(* IEC 61131-3 sources: daoli-st-library/DL_Process (part 47) *)

(* ---- FB_DL_QuarterCellCutSeq.st ---- *)
(*
  FB_DL_QuarterCellCutSeq  —  极片分切顺控（刀轴相位 + 张力窗 + 废边回收） / Electrode slitting sequencer with blade phase, tension window and trim recovery
  分类 Category : DL_Process
  版本 Version  : 1.0.0
  来源 Source   : roadmap-li-p2 — 锂电极片分切工站真缺口
  溯源 Origin   : 道莅 clean-room 实现；刀轴相位对齐 + 张力窗监督 + 废边回收联锁为公开分切工艺逻辑，未复制任何源码行
  功能 Function : 1) 三段顺控：ePhase 刀轴相位对齐（fBladePhaseDeg 进目标容差带）→
                  eRun 分切运行（张力窗 fTensionN 双向监督 + 废边回收信号 bTrimOk 监督）→
                  eStop 收料停机（tStop 到时）→ eDone；2) 相位对齐超时保护；
                  3) 故障级单码 03A0，归因由 eCause 独立成员承载（R190）；
                  4) 信息级 04C8 = 分切循环完成沿；5) 解除式全当拍量（R240）。
  接口 Interface: 输入相位/张力/废边信号与复位位；输出状态/相位镜像/张力窗镜像/码
  边界 Boundary : ① 组态闸：fPhaseTolDeg <= 0.0、fTensionHiN <= fTensionLoN、tPhaseTmo <= T#0S、
                  tStop <= T#0S → 03A0 锁存；② 相位判据为双向容差式，相位量纲约定
                  0~360 单调注入（跨零归一由调用方完成，本件不内联 MOD 以免非标准扩展）；
                  ③ 浮点禁 = / <> 判等；④ 全部 TON / R_TRIG 段 0 无条件周期调用；
                  ⑤ 故障相迁出唯一路径 = bReset 上升沿；⑥ 零全局耦合（无 GVL / %I %Q %M）。
  依赖 Depends  : Standard.library（TON / R_TRIG）
  码表 Error codes（Process 段 0005，故障窗口 03A0 / 信息窗口 04C8）:
    16#0005_03A0 故障级：分切故障总码（组态非法 / 相位对齐超时 / 张力越窗 / 废边回收异常），
                 锁存至 bReset 上升沿；归因见 eCause，不新增码位（派单硬约束单码）
    16#0005_04C8 信息级：分切循环完成沿（收料停机完成进 eDone 单拍）
  修订历史 Revision :
    2026-11-19  v1.0.0  R43 首版（批次 1 · 序号 4）
*)

TYPE E_DL_QcsState :
(
    eIdle  := 0,      // 未使能待启动 / Idle, waiting start
    ePhase := 10,     // 刀轴相位对齐中 / Blade phase alignment
    eRun   := 20,     // 分切运行（张力窗 + 废边监督） / Slitting under tension and trim supervision
    eStop  := 30,     // 收料停机中 / Web stop
    eDone  := 50,     // 循环完成 / Done
    eFault := 90      // 故障锁存相 / Fault latched phase
);
END_TYPE

TYPE E_DL_QcsCause :
(
    eNone       := 0, // 无故障成因 / No cause
    eCfgIllegal := 1, // 组态非法 / Illegal configuration
    ePhaseTmo   := 2, // 相位对齐超时 / Phase alignment timeout
    eTensionDev := 3, // 张力越窗 / Tension out of window
    eTrimLost   := 4  // 废边回收异常 / Trim recovery lost
);
END_TYPE

FUNCTION_BLOCK FB_DL_QuarterCellCutSeq
VAR_INPUT
    fBladePhaseDeg  : REAL := 0.0;       // 刀轴实测相位 [°]，0~360 单调注入 / Blade shaft phase
    fPhaseTgtDeg    : REAL := 90.0;      // 目标相位 [°] / Target phase
    fPhaseTolDeg    : REAL := 1.0;       // 相位容差带 [°]，域 > 0 / Phase tolerance
    fTensionN       : REAL := 0.0;       // 实测极片张力 [N] / Measured web tension
    fTensionLoN     : REAL := 20.0;      // 张力窗下限 [N] / Tension low limit
    fTensionHiN     : REAL := 60.0;      // 张力窗上限 [N] / Tension high limit
    bTrimOk         : BOOL := FALSE;     // 废边回收正常信号（电平）[-] / Trim recovery healthy
    tPhaseTmo       : TIME := T#5S;      // 相位对齐超时 [ms]，域 > 0 / Phase timeout
    tStop           : TIME := T#2S;      // 收料停机时长 [ms]，域 > 0 / Web stop duration
    bStart          : BOOL := FALSE;     // 启动命令（电平）[-] / Start command
    bReset          : BOOL := FALSE;     // 复位命令，上升沿清故障 [-] / Reset edge
END_VAR
VAR_OUTPUT
    eState          : E_DL_QcsState;     // 状态出口，段 6 单点映射 / State outlet
    eCause          : E_DL_QcsCause;     // 故障成因出口（R190） / Fault cause outlet
    fPhaseDegOut    : REAL;              // 相位镜像 [°] / Phase mirror
    bPhaseOk        : BOOL;              // 相位达窗镜像 [-] / Phase in-window mirror
    bTensionOk      : BOOL;              // 张力在窗镜像 [-] / Tension in-window mirror
    bCycleDone      : BOOL;              // 循环完成标志 [-] / Cycle done flag
    bError          : BOOL;              // 故障锁存标志 [-] / Fault latch flag
    nErrId          : UDINT;             // 事件码，0 = 无事件 / Event code
END_VAR
VAR
    _eState         : E_DL_QcsState := E_DL_QcsState.eIdle;   // 内部相位（CASE 唯一写入目标） / Internal phase
    _eCause         : E_DL_QcsCause := E_DL_QcsCause.eNone;   // 故障成因锁存（锁存量） / Latched cause
    tonPhase        : TON;               // 相位对齐计时，每周期无条件调用 / Phase timer
    tonStop         : TON;               // 收料停机计时，每周期无条件调用 / Stop timer
    rtReset         : R_TRIG;            // 复位沿实例，每周期无条件调用 / Reset edge
    _bPhaseOk       : BOOL;              // 相位达窗当拍量 [-] / Phase verdict
    _bTensionOk     : BOOL;              // 张力在窗当拍量 [-] / Tension verdict
    _bCfgBad        : BOOL;              // 组态非法当拍量 [-] / Config illegal
    _bFault         : BOOL;              // 故障锁存位（锁存量） / Latched fault bit
    _uFault         : UDINT;             // 故障码锁存（锁存量） / Latched fault code
    _uInfo          : UDINT;             // 信息码，每拍重算 / Transient info code
END_VAR

(* —— 段 0：沿实例与定时器无条件周期刷新 —— *)
_bPhaseOk := ABS(fBladePhaseDeg - fPhaseTgtDeg) <= fPhaseTolDeg;                 // 相位容差判据 / Phase tolerance verdict
_bTensionOk := (fTensionN >= fTensionLoN - 1.0E-6) AND (fTensionN <= fTensionHiN + 1.0E-6);  // 张力容差窗 / Tension window verdict
_bCfgBad := (fPhaseTolDeg <= 0.0) OR (fTensionHiN <= fTensionLoN)
            OR (tPhaseTmo <= T#0S) OR (tStop <= T#0S);                          // 组态非法当拍量 / Config illegal
rtReset(CLK := bReset);                                                        // 复位沿，每拍必调 / Reset edge
tonPhase(IN := (_eState = E_DL_QcsState.ePhase), PT := tPhaseTmo);             // 相位对齐计时 / Phase timer
tonStop(IN := (_eState = E_DL_QcsState.eStop), PT := tStop);                   // 收料停机计时 / Stop timer

(* —— 段 1：单拍量预清零（锁存量不入清单） —— *)
_uInfo := 16#0000_0000;            // 信息码每拍重算 / Info recomputed
fPhaseDegOut := 0.0;               // 相位镜像缺省 0 / Phase mirror default
bPhaseOk := FALSE;                 // 相位镜像缺省 FALSE / Phase flag default
bTensionOk := FALSE;               // 张力镜像缺省 FALSE / Tension flag default
bCycleDone := FALSE;               // 完成标志缺省 FALSE / Done default
nErrId := 16#0000_0000;            // 事件码缺省无事件 / Event code default

(* —— 段 2：复位沿 + 组态域闸 —— *)
IF rtReset.Q THEN                              // rtReset.Q = 当拍量 / current scan
    _bFault := FALSE;                          // 清故障锁存位（锁存量） / Clear fault latch
    _uFault := 16#0000_0000;                   // 清故障锁存码（锁存量） / Clear fault code
    _eCause := E_DL_QcsCause.eNone;            // 清成因（锁存量） / Clear cause
    IF _eState = E_DL_QcsState.eFault THEN
        _eState := E_DL_QcsState.eIdle;        // 故障相迁出：回未使能 / Fault exit to idle
    END_IF
END_IF
IF _bCfgBad THEN                               // 组态域闸 / Config gate
    _uFault := 16#0005_03A0;                   // 故障级：分切故障总码 / Process fault code
    _eCause := E_DL_QcsCause.eCfgIllegal;      // 归因：组态非法 / Cause: illegal config
    _bFault := TRUE;                           // 标志与码位配对（R45） / Flag paired with code
END_IF

(* —— 段 3：超时 / 张力越窗 / 废边异常（判据当拍量） —— *)
IF (NOT _bFault) AND tonPhase.Q THEN           // 相位对齐超时 / Phase timeout
    _uFault := 16#0005_03A0;
    _eCause := E_DL_QcsCause.ePhaseTmo;        // 归因：相位超时 / Cause: phase timeout
    _bFault := TRUE;
END_IF
IF (NOT _bFault) AND (_eState = E_DL_QcsState.eRun) AND (NOT _bTensionOk) THEN   // 运行期张力越窗 / Tension deviation
    _uFault := 16#0005_03A0;
    _eCause := E_DL_QcsCause.eTensionDev;      // 归因：张力越窗 / Cause: tension
    _bFault := TRUE;
END_IF
IF (NOT _bFault) AND (_eState = E_DL_QcsState.eRun) AND (NOT bTrimOk) THEN       // 废边回收异常 / Trim lost
    _uFault := 16#0005_03A0;
    _eCause := E_DL_QcsCause.eTrimLost;        // 归因：废边异常 / Cause: trim lost
    _bFault := TRUE;
END_IF

(* —— 段 4：故障解除式（R240；全当拍量）：rtReset.Q / NOT _bCfgBad / NOT tonPhase.Q —— *)
IF rtReset.Q AND (NOT _bCfgBad) AND (NOT tonPhase.Q) THEN
    _bFault := FALSE;                          // 清故障锁存位（锁存量） / Clear fault latch
    _uFault := 16#0000_0000;                   // 清故障锁存码（锁存量） / Clear fault code
    _eCause := E_DL_QcsCause.eNone;            // 清成因（锁存量） / Clear cause
END_IF

(* —— 段 4A：故障锁存相位迁移闸 —— *)
IF _bFault AND (_eState <> E_DL_QcsState.eFault) THEN
    _eState := E_DL_QcsState.eFault;           // 锁存即入故障相 / Latch enters fault phase
END_IF

(* —— 段 5：相位机（CASE 全覆盖 + ELSE 兜底） —— *)
CASE _eState OF

E_DL_QcsState.eIdle:
    IF bStart AND (NOT _bFault) THEN           // 启动条件 / Start gate
        _eState := E_DL_QcsState.ePhase;       // 进相位对齐相 / Enter phase alignment
    END_IF

E_DL_QcsState.ePhase:
    IF _bPhaseOk THEN                          // 出口 1：相位达窗 / Phase reached
        _eState := E_DL_QcsState.eRun;         // 进分切运行相 / Enter slitting
    ELSIF NOT bStart THEN                      // 出口 2：撤启动（R98 双出口） / Start released
        _eState := E_DL_QcsState.eIdle;        // 回未使能 / Back to idle
    END_IF

E_DL_QcsState.eRun:
    IF NOT bStart THEN                         // 撤启动：进停机相 / Start released enters stop
        _eState := E_DL_QcsState.eStop;
    END_IF

E_DL_QcsState.eStop:
    IF tonStop.Q THEN                          // 停机计时到 / Stop elapsed
        _uInfo := 16#0005_04C8;                // 信息级：循环完成沿 / Info: cycle complete edge
        _eState := E_DL_QcsState.eDone;        // 进完成相 / Enter done
    END_IF

E_DL_QcsState.eDone:
    IF bStart THEN                             // 新循环请求 / New cycle request
        _eState := E_DL_QcsState.ePhase;       // 进相位相 / Enter phase
    END_IF

E_DL_QcsState.eFault:
    ;                                          // 故障相：仅段 4 复位沿可迁出 / Only reset exits

ELSE
    _uFault := 16#0005_03A0;                   // 故障级：非法相位兜底（归并总码） / Illegal phase fallback
    _eCause := E_DL_QcsCause.eCfgIllegal;      // 归因：相位非法归并组态 / Cause: phase illegal
    _bFault := TRUE;
    _eState := E_DL_QcsState.eFault;           // 强制回故障相 / Force fault phase

END_CASE

(* —— 段 6：出口单点映射（名实同源；锁存码回放） —— *)
fPhaseDegOut := fBladePhaseDeg;                    // 相位镜像 / Phase mirror
bPhaseOk := _bPhaseOk AND (NOT _bFault);           // 相位达窗镜像 / Phase mirror
bTensionOk := _bTensionOk AND (NOT _bFault);       // 张力窗镜像 / Tension mirror
bCycleDone := (_eState = E_DL_QcsState.eDone);     // 完成标志 / Done flag
IF _bFault THEN
    nErrId := _uFault;                         // 故障锁存码回放 / Replay latched code
ELSE
    nErrId := _uInfo;                          // 信息码 / Transient info
END_IF
bError := _bFault;                             // 故障标志同源 / Flag from latch
eState := _eState;                             // 状态出口 / State outlet
eCause := _eCause;                             // 成因出口 / Cause outlet

END_FUNCTION_BLOCK

(* ---- FB_DL_QuenchTemperLineSeq.st ---- *)
(*==============================================================================
  Component : FB_DL_QuenchTemperLineSeq
  Category  : DL_Process
  Type      : FB
  Complexity: C4
  VERSION   : v1.0.0
  功能      : 淬火-回火联动线全流程顺控（上料/加热/保温/淬火/沥液/回火/冷却/下料）
  开源溯源  : 道莅原创 clean-room 自研（无外部代码引用）｜License: MIT
  边界条件  : ① 本件只编排相与时序闸，不驱动阀门接触器；执行器由 IO 映射层按相指示位驱动。
              ② E1 仅加热相与沥液相可重试（定时器自复位后重新计时），预算 nRetryMax 耗尽升 E2。
              ③ E3 判据（急停断开 / 安全门未闭 / 液位低于下限 / 介质超温）同拍置 bSafeCut；
                 锁存解除唯一路径 = bReset 沿且安全条件已恢复（R152），bStop 不清 E3。
              ④ 配比约束（R100）：atPhaseTmo[1] 加热窗须宽于实测升温时间；atPhaseTmo[6] 回火总窗
                 须 ≥ 升温 + 保温整定之和，否则回火带内判据永不到时。
              ⑤ 复位作用域（R311）：bReset 沿清 E2/E3 锁存 + 节拍累加 + 重试计数；bStop 只清 E2 与相位。
              ⑥ 默认引脚组合自证（R114）：握手类（bPartLoaded / bUnloadPermit / bDrained /
                 bQuenchImmersion）默认 FALSE，默认组合无法越过任一握手直达完成相；使能类（bDoorClosed /
                 bEStopHealthy）默认 TRUE 与 bEnable 同族，断线由硬件安全回路保证，不靠软件默认值兜底。
  状态机    : eIdle 待机 / eLoad 上料 / eHeat 加热 / eSoak 保温 / eQuench 淬火 / eDrain 沥液 /
              eTemper 回火 / eCool 冷却 / eUnload 下料 / eFault 故障停(E2) / eSafeStop 安全断能(E3)
  自检      : R1 零 GVL ｜ R2 零物理地址 ｜ R3 纯 IEC 61131-3 ｜ R4 非有限自反判 + 除零先判 ｜
              R6 CASE 含 ELSE ｜ R7 八 TON 两沿段 0 无条件刷新 ｜ R10 仅标准转换函数 ｜ R14 无属性件
==============================================================================*)
TYPE E_DL_QtlPhase :
(
    eIdle     := 0,     (* 待机：等启动沿 / Idle, waiting for start edge *)
    eLoad     := 10,    (* 上料相：等上料到位 / Loading, wait load-in-position *)
    eHeat     := 20,    (* 加热相：升到保温带（E1 可重试）/ Heating, retryable *)
    eSoak     := 30,    (* 保温相：保温到时 / Soaking *)
    eQuench   := 40,    (* 淬火相：浸没且到时 / Quenching, immersed and timed *)
    eDrain    := 50,    (* 沥液相：等回液到位（E1 可重试）/ Draining, retryable *)
    eTemper   := 60,    (* 回火相：带内且总窗到时 / Tempering, in band and window *)
    eCool     := 70,    (* 冷却相：空冷到出料温度 / Cooling to unload temperature *)
    eUnload   := 80,    (* 下料相：等下料允许 / Unloading, wait permit *)
    eFault    := 90,    (* 故障停待复位（E2）/ Fault stop awaiting reset, E2 *)
    eSafeStop := 95     (* 安全侧断能（E3）/ Safety energy cut, E3 *)
);
END_TYPE
TYPE E_DL_QtlCause :
(
    eNone      := 0,    (* 无异常 / No anomaly *)
    eLoadTmo   := 1,    (* 上料超时 / Load timeout *)
    eHeatTmo   := 2,    (* 加热超时（E1 记录后重试）/ Heat timeout, retried *)
    eSoakTmo   := 3,    (* 保温超时 / Soak timeout *)
    eQuenchTmo := 4,    (* 淬火到时未浸没 / Quench timed out without immersion *)
    eDrainTmo  := 5,    (* 沥液超时（E1 记录后重试）/ Drain timeout, retried *)
    eTemperTmo := 6,    (* 回火超时（带内未达）/ Tempering timeout *)
    eCoolTmo   := 7,    (* 冷却超时 / Cooling timeout *)
    eUnloadTmo := 8,    (* 下料超时 / Unload timeout *)
    eRetryOver := 9,    (* 重试预算耗尽（E1 升 E2）/ Retry budget exhausted *)
    eSigBad    := 10,   (* 工件温度信号非有限（E2）/ Part temperature non-finite *)
    eEstopOpen := 11,   (* 急停回路断开（E3）/ E-stop circuit open *)
    eDoorOpen  := 12,   (* 安全门未闭合（E3）/ Guard door open *)
    eLevelLow  := 13,   (* 淬火槽液位低于下限（E3）/ Bath level low *)
    eMediumHi  := 14,   (* 淬火介质超温（E3）/ Medium over-temperature *)
    eCfgBad    := 15,   (* 组态非法（E2）/ Illegal configuration *)
    ePhaseBad  := 16    (* 非法相位兜底（E2）/ Illegal phase fallback *)
);
END_TYPE
TYPE E_DL_QtlGrade :
(
    eG0 := 0,           (* 无异常 / No anomaly *)
    eG1 := 1,           (* E1 可恢复重试：记录后重试，不置 bError / E1 retried, recorded only *)
    eG2 := 2,           (* E2 停机待复位 / E2 stop, awaiting reset *)
    eG3 := 3            (* E3 安全侧立即断能 / E3 immediate safety energy cut *)
);
END_TYPE

FUNCTION_BLOCK FB_DL_QuenchTemperLineSeq
VAR_INPUT
    bStart        : BOOL := FALSE;      (* 启动沿（eIdle 入 eLoad） [-] / Start rising edge *)
    bStop         : BOOL := FALSE;      (* 中止：回 eIdle 并清 E2 锁存（不清 E3） [-] / Abort, clears E2 only *)
    bReset        : BOOL := FALSE;      (* 复位沿：清全部锁存 + 节拍 + 重试（R311） [-] / Reset edge *)
    bPartLoaded   : BOOL := FALSE;      (* 上料到位（默认 FALSE 禁跳步） [-] / Load in position *)
    bUnloadPermit : BOOL := FALSE;      (* 下料允许（默认 FALSE 禁跳步） [-] / Unload permit *)
    bQuenchOil    : BOOL := TRUE;       (* 介质：TRUE 油淬 / FALSE 水淬 [-] / Oil when TRUE *)
    bQuenchImmersion : BOOL := FALSE;   (* 淬火浸没到位（默认 FALSE 禁跳步） [-] / Quench immersion OK *)
    bDrained      : BOOL := FALSE;      (* 沥液回液到位（默认 FALSE 禁跳步） [-] / Drain back complete *)
    bDoorClosed   : BOOL := TRUE;       (* 安全门闭合（使能类引脚，默认 TRUE） [-] / Guard door closed *)
    bEStopHealthy : BOOL := TRUE;       (* 急停回路正常（使能类引脚，默认 TRUE） [-] / E-stop healthy *)
    fMediumTempC  : LREAL := 0.0;       (* 淬火介质温度实测 [℃] / Medium temperature [degC] *)
    fLevelPct     : LREAL := 0.0;       (* 淬火槽液位实测 [%] / Bath level [%] *)
    fPartTempC    : LREAL := 0.0;       (* 工件温度实测（升温与冷却判据） [℃] / Part temperature [degC] *)
    fSoakSetC     : LREAL := 850.0;     (* 保温设定温度，域 > 0 [℃] / Soak setpoint [degC] *)
    fTemperSetC   : LREAL := 550.0;     (* 回火设定温度，域 > 0 [℃] / Temper setpoint [degC] *)
    fSoakTolC     : LREAL := 15.0;      (* 保温与回火带共用半宽，域 > 0 [℃] / Band half-width [degC] *)
    fMediumMaxC   : LREAL := 60.0;      (* 介质温度上限，域 > 0（E3 判据） [℃] / Medium limit [degC] *)
    fLevelMinPct  : LREAL := 70.0;      (* 液位安全下限，域 0..100（E3 判据） [%] / Level floor [%] *)
    fCoolSetC     : LREAL := 80.0;      (* 冷却出料温度上限，域 > 0 [℃] / Cool-down unload limit [degC] *)
    atPhaseTmo    : ARRAY[0..8] OF TIME := [T#3M, T#45M, T#90M, T#15M, T#8M, T#3M, T#120M, T#30M, T#3M];   (* 超时窗 [ms]，下标 0..8 = 上料/加热/保温/油淬/水淬/沥液/回火/冷却/下料 / Phase windows [ms] *)
    nRetryMax     : UINT := 2;          (* 单相 E1 重试预算，域 1..9（0 入组态闸） [次] / Retry budget *)
    fCycleSec     : LREAL := 0.0;       (* 扫描周期（<=0 用缺省 0.01s） [s] / Scan cycle [s] *)
END_VAR
VAR_OUTPUT
    eState        : E_DL_QtlPhase;      (* 当前相（HMI 诊断） [-] / Present phase *)
    eCause        : E_DL_QtlCause;      (* 成因（锁存回放，R189） [-] / Latched cause playback *)
    eGrade        : E_DL_QtlGrade;      (* 异常分级出口 [-] / Exception grade outlet *)
    bError        : BOOL;               (* 故障标志（E2/E3 为 TRUE，E1 不置） [-] / Error flag *)
    bSafeCut      : BOOL;               (* 安全侧断能指令（E3 常 TRUE 至复位） [-] / Safety energy cut *)
    bHeatActive   : BOOL;               (* 加热相指示（供 IO 层驱动加热阀） [-] / Heating indicator *)
    bQuenchActive : BOOL;               (* 淬火相指示（供 IO 层驱动淬火机构） [-] / Quench indicator *)
    bDone         : BOOL;               (* 单拍完成脉冲 [-] / One-scan done pulse *)
    nPieceCount   : UDINT;              (* 累计产量（饱和于 UDINT 上限） [件] / Piece count, saturating *)
    tCycleLast    : TIME;               (* 最近一件节拍 [ms] / Last piece cycle [ms] *)
    fCycleAvgS    : LREAL;              (* 平均节拍（无件输出 0） [s] / Average cycle [s] *)
    nRetryUsed    : UINT;               (* 当前相已用重试次数 [次] / Retries used in phase *)
END_VAR
VAR
    _ePhase      : E_DL_QtlPhase := E_DL_QtlPhase.eIdle;    (* 内部相（CASE 唯一写入目标） [-] / Internal phase *)
    _ePhasePrev  : E_DL_QtlPhase := E_DL_QtlPhase.eIdle;    (* 上拍相快照（相迁移后置用） [-] / Previous phase *)
    _eCause      : E_DL_QtlCause := E_DL_QtlCause.eNone;    (* 成因锁存量 [-] / Latched cause *)
    _eGrade      : E_DL_QtlGrade := E_DL_QtlGrade.eG0;      (* 分级锁存量 [-] / Latched grade *)
    _bFault      : BOOL := FALSE;       (* E2 锁存位（解除 = bReset 沿或 bStop） [-] / E2 latch *)
    _bSafeLatch  : BOOL := FALSE;       (* E3 锁存位（解除 = bReset 沿且安全恢复） [-] / E3 latch *)
    _bFaultReq   : BOOL := FALSE;       (* 单拍故障请求（段 1 预清，段 6 落地） [-] / One-scan fault request *)
    _bDonePulse  : BOOL := FALSE;       (* 单拍完成标志（段 1 预清） [-] / One-scan done flag *)
    _bMediumBad  : BOOL := FALSE;       (* 介质温度非有限或超上限 [-] / Medium bad *)
    _bLevelBad   : BOOL := FALSE;       (* 液位非有限或低于下限 [-] / Level bad *)
    _bPartBad    : BOOL := FALSE;       (* 工件温度非有限 [-] / Part temperature non-finite *)
    _bSoakBand   : BOOL := FALSE;       (* 保温带内判据 [-] / In soak band *)
    _bTemperBand : BOOL := FALSE;       (* 回火带内判据 [-] / In temper band *)
    _bCfgBad     : BOOL := FALSE;       (* 组态非法当拍量 [-] / Configuration bad *)
    _nRetry      : UINT := 0;           (* 当前相重试计数（相迁移后置清） [次] / Retry counter *)
    _nPiece      : UDINT := 0;          (* 产量累计锁存（饱和） [件] / Piece count latch *)
    _nIdx        : INT := 0;            (* 相窗遍历索引（循环变量） [-] / Loop index *)
    _fCycleAccS  : LREAL := 0.0;        (* 本件节拍累加 [s] / Cycle accumulator *)
    _fCycleSumS  : LREAL := 0.0;        (* 节拍总和（均值分子） [s] / Cycle sum *)
    _fCy         : LREAL := 0.0;        (* 当拍有效周期 [s] / Effective cycle *)
    _tCycleLast  : TIME := T#0S;        (* 最近节拍锁存 [ms] / Last cycle latch *)
    _tQuenchTmo  : TIME := T#15M;       (* 当拍淬火窗（按介质选择） [ms] / Active quench window [ms] *)
    tonLoad      : TON;                 (* 上料超时（段 0 无条件调用） / Load timeout *)
    tonHeat      : TON;                 (* 加热超时（自复位，E1 可重试） / Heat timeout, self-reset *)
    tonSoak      : TON;                 (* 保温超时 / Soak timeout *)
    tonQuench    : TON;                 (* 淬火超时（按介质选窗） / Quench timeout *)
    tonDrain     : TON;                 (* 沥液超时（自复位，E1 可重试） / Drain timeout, self-reset *)
    tonTemper    : TON;                 (* 回火总窗（升温 + 保温） / Temper total window *)
    tonCool      : TON;                 (* 冷却超时 / Cool timeout *)
    tonUnload    : TON;                 (* 下料超时 / Unload timeout *)
    rtStart      : R_TRIG;              (* 启动沿（段 0 无条件调用） / Start edge *)
    rtReset      : R_TRIG;              (* 复位沿（段 0 无条件调用） / Reset edge *)
END_VAR
VAR CONSTANT
    DL_QTL_CYDEF    : LREAL := 0.01;        (* 缺省扫描周期 [s] / Default scan cycle [s] *)
    DL_QTL_PCMAX    : UDINT := 4294967295;  (* 产量计数饱和上限 [件] / Piece count ceiling *)
    DL_QTL_RETRYTOP : UINT := 9;            (* 重试预算可配域顶 [次] / Retry configurable ceiling *)
    DL_QTL_PCTOP    : LREAL := 100.0;       (* 液位百分比满量程 [%] / Level full scale [%] *)
END_VAR

(*-----------------------------------------------------------------------------
  方法 ResetFault：清 E2/E3 锁存（唯一解除入口，R152 可达性自证）
  契约：入参 bSafetyOk 表示安全条件已恢复；返回 TRUE = 本次确实清除了锁存。
  E2 恒可清；E3 仅当 bSafetyOk 为 TRUE 才可清（否则锁存保持，解除路径显式可达）。
  作用域：清 _bFault / _bSafeLatch / _eCause / _eGrade / _nRetry，并把相位迁回 eIdle。
-----------------------------------------------------------------------------*)
METHOD PUBLIC ResetFault : BOOL
VAR_INPUT
    bSafetyOk : BOOL := FALSE;      (* 安全条件已恢复（E3 解除前置） [-] / Safety conditions recovered *)
END_VAR
VAR
    _bCleared : BOOL := FALSE;      (* 本次是否清除过锁存 [-] / Cleared this call *)
END_VAR

ResetFault := FALSE;                (* 返回预置安全值 / Preset safe return *)
_bCleared := FALSE;
IF _bSafeLatch THEN
    IF bSafetyOk THEN
        _bSafeLatch := FALSE;       (* E3 解除：安全侧恢复后允许 / E3 released after safety recovery *)
        _bCleared := TRUE;
    END_IF
ELSIF _bFault THEN
    _bFault := FALSE;               (* E2 解除：无条件可清 / E2 released unconditionally *)
    _bCleared := TRUE;
END_IF
IF _bCleared THEN
    _eCause := E_DL_QtlCause.eNone;     (* 清成因 / Clear cause *)
    _eGrade := E_DL_QtlGrade.eG0;       (* 清分级 / Clear grade *)
    _nRetry := 0;                       (* 清重试预算占用 / Clear retry usage *)
    _ePhase := E_DL_QtlPhase.eIdle;     (* 迁回待机 / Back to idle *)
END_IF
ResetFault := _bCleared;            (* 真值返回 / Final return *)
END_METHOD

(*-----------------------------------------------------------------------------
  方法 CalcCycleTime：本件节拍换算（毫秒取整 + 双向域闸，无跨周期驻留）
  口径：NaN 自反检出 -> 返回哨兵零点 T#0S（还原方向不饱和，R81）；
        Inf 用差值自减检出 -> 亦返回哨兵零点；负值拒收；
        超 TIME 可表上限先钳后转（R153 取整前实数上限兜底）。
-----------------------------------------------------------------------------*)
METHOD PUBLIC CalcCycleTime : TIME
VAR
    fMs   : LREAL := 0.0;           (* 节拍毫秒暂存 [ms] / Milliseconds scratch *)
    fMsCl : LREAL := 0.0;           (* 钳位后毫秒 [ms] / Clamped milliseconds *)
    diMs  : DINT := 0;              (* 整型毫秒（钳位后转换，防溢出翻转） [ms] / Integer milliseconds *)
END_VAR

CalcCycleTime := T#0S;              (* 哨兵零点 / Sentinel zero *)
fMs := _fCycleAccS * 1000.0;        (* 秒 -> 毫秒 [ms] / Second to millisecond *)
IF (fMs <> fMs) OR ((fMs - fMs) <> (fMs - fMs)) OR (fMs < 0.0) THEN
    CalcCycleTime := T#0S;          (* 域闸：NaN 自反 / Inf 差值自减 / 负值，均拒收 / Domain gate *)
    RETURN;
END_IF
IF fMs > 2147483647.0 THEN
    fMsCl := 2147483647.0;          (* 先钳到 TIME 可表毫秒上限 / Clamp to TIME ceiling *)
ELSE
    fMsCl := fMs;
END_IF
diMs := LREAL_TO_DINT(fMsCl);       (* 钳位后整型转换（R10 标准函数） / Clamped integer conversion *)
CalcCycleTime := DINT_TO_TIME(diMs);(* 标准转换链 / Standard conversion chain *)
END_METHOD

(* —— 段 0：三模拟量非有限判定 + 组态闸 + 淬火窗选择 + 周期派生 + 八 TON 两沿无条件刷新（R7） —— *)
_bMediumBad := (fMediumTempC <> fMediumTempC)
            OR ((fMediumTempC - fMediumTempC) <> (fMediumTempC - fMediumTempC))
            OR (fMediumTempC > fMediumMaxC);      (* NaN 自反 + Inf 差值 + 超上限 / NaN, Inf, over-limit *)
_bLevelBad := (fLevelPct <> fLevelPct)
           OR ((fLevelPct - fLevelPct) <> (fLevelPct - fLevelPct))
           OR (fLevelPct < fLevelMinPct);         (* NaN 自反 + Inf 差值 + 低于下限 / NaN, Inf, low level *)
_bPartBad := (fPartTempC <> fPartTempC)
          OR ((fPartTempC - fPartTempC) <> (fPartTempC - fPartTempC));   (* 工件温度非有限 / Part temp non-finite *)
_bCfgBad := (nRetryMax = 0) OR (nRetryMax > DL_QTL_RETRYTOP)
         OR (fSoakSetC <= 0.0) OR (fTemperSetC <= 0.0) OR (fSoakTolC <= 0.0)
         OR (fMediumMaxC <= 0.0) OR (fCoolSetC <= 0.0)
         OR (fLevelMinPct < 0.0) OR (fLevelMinPct > DL_QTL_PCTOP);   (* 静态组态域闸全枚举 / Static config gate *)
FOR _nIdx := 0 TO 8 DO
    IF atPhaseTmo[_nIdx] <= T#0S THEN
        _bCfgBad := TRUE;                          (* 任一相窗非正 -> 组态非法 / Non-positive phase window *)
    END_IF
END_FOR
IF bQuenchOil THEN
    _tQuenchTmo := atPhaseTmo[3];                  (* 油淬窗 / Oil quench window *)
ELSE
    _tQuenchTmo := atPhaseTmo[4];                  (* 水淬窗 / Water quench window *)
END_IF
IF fCycleSec > 0.0 THEN
    _fCy := fCycleSec;                             (* 组态周期有效 / Configured cycle valid *)
ELSE
    _fCy := DL_QTL_CYDEF;                          (* 周期缺省兜底 / Default cycle *)
END_IF
_bSoakBand := (NOT _bPartBad) AND (ABS(fPartTempC - fSoakSetC) <= fSoakTolC);     (* 保温带内（容差比较） / In soak band *)
_bTemperBand := (NOT _bPartBad) AND (ABS(fPartTempC - fTemperSetC) <= fSoakTolC); (* 回火带内（共用半宽） / In temper band *)
rtStart(CLK := bStart);                            (* 启动沿，每拍必调 / Start edge every scan *)
rtReset(CLK := bReset);                            (* 复位沿，每拍必调 / Reset edge every scan *)
tonLoad(IN := (_ePhase = E_DL_QtlPhase.eLoad), PT := atPhaseTmo[0]);              (* 上料超时 / Load window *)
tonHeat(IN := (_ePhase = E_DL_QtlPhase.eHeat) AND (NOT tonHeat.Q), PT := atPhaseTmo[1]);   (* 加热自复位窗（R188） / Heat self-reset *)
tonSoak(IN := (_ePhase = E_DL_QtlPhase.eSoak), PT := atPhaseTmo[2]);              (* 保温超时 / Soak window *)
tonQuench(IN := (_ePhase = E_DL_QtlPhase.eQuench), PT := _tQuenchTmo);            (* 淬火超时 / Quench window *)
tonDrain(IN := (_ePhase = E_DL_QtlPhase.eDrain) AND (NOT tonDrain.Q), PT := atPhaseTmo[5]); (* 沥液自复位窗 / Drain self-reset *)
tonTemper(IN := (_ePhase = E_DL_QtlPhase.eTemper), PT := atPhaseTmo[6]);          (* 回火总窗 / Temper window *)
tonCool(IN := (_ePhase = E_DL_QtlPhase.eCool), PT := atPhaseTmo[7]);              (* 冷却超时 / Cool window *)
tonUnload(IN := (_ePhase = E_DL_QtlPhase.eUnload), PT := atPhaseTmo[8]);          (* 下料超时 / Unload window *)

(* —— 段 1：单拍量预清零（不含锁存/累加/快照量，R107）+ 相迁移后置 —— *)
_bFaultReq := FALSE;                               (* 单拍故障请求预清 / Fault request preset *)
_bDonePulse := FALSE;                              (* 单拍完成标志预清 / Done pulse preset *)
bError := FALSE;                                   (* 故障标志预清（出口 OR 汇总） / Error preset *)
IF _ePhase <> _ePhasePrev THEN
    _nRetry := 0;                                  (* 相迁移：重试预算复位 / Phase change: retry reset *)
    IF _eGrade = E_DL_QtlGrade.eG1 THEN
        _eGrade := E_DL_QtlGrade.eG0;              (* E1 记录随相推进清零（信息级可重算） / E1 cleared on advance *)
        _eCause := E_DL_QtlCause.eNone;
    END_IF
END_IF

(* —— 段 2：E3 安全侧拦截（最高优先级，同拍断能 + 归因唯一 + 迁相） —— *)
IF (NOT bEStopHealthy) OR (NOT bDoorClosed) OR _bLevelBad OR _bMediumBad THEN
    IF NOT _bSafeLatch THEN
        _bSafeLatch := TRUE;                       (* 锁存 / Latch *)
        _eGrade := E_DL_QtlGrade.eG3;              (* 分级 E3 / Grade E3 *)
        bError := TRUE;                            (* 分级标志同段置位（R45 配对） / Error pairing *)
        IF NOT bEStopHealthy THEN
            _eCause := E_DL_QtlCause.eEstopOpen;   (* 归因：急停断开 / Cause: E-stop *)
        ELSIF NOT bDoorClosed THEN
            _eCause := E_DL_QtlCause.eDoorOpen;    (* 归因：安全门未闭 / Cause: door *)
        ELSIF _bLevelBad THEN
            _eCause := E_DL_QtlCause.eLevelLow;    (* 归因：液位低 / Cause: level *)
        ELSE
            _eCause := E_DL_QtlCause.eMediumHi;    (* 归因：介质超温 / Cause: medium *)
        END_IF
    END_IF
    _ePhase := E_DL_QtlPhase.eSafeStop;            (* 同步迁安全相 / Migrate to safety stop *)
END_IF

(* —— 段 3：组态闸入 E2（E3 优先，安全相内不重复置因） —— *)
IF _bCfgBad AND (NOT _bSafeLatch) AND (NOT _bFault) THEN
    _bFault := TRUE;                               (* E2 锁存 / Latch E2 *)
    _eGrade := E_DL_QtlGrade.eG2;                  (* 分级 E2 / Grade E2 *)
    _eCause := E_DL_QtlCause.eCfgBad;              (* 归因：组态非法 / Cause: config *)
    _ePhase := E_DL_QtlPhase.eFault;               (* 同步迁相（R252） / Migrate *)
END_IF

(* —— 段 4：迁出链（复位沿 > 中止；作用域逐项声明 R311） —— *)
IF rtReset.Q THEN
    _bFault := FALSE;                              (* 作用域①：清 E2 锁存 / Clear E2 *)
    IF NOT ((NOT bEStopHealthy) OR (NOT bDoorClosed) OR _bLevelBad OR _bMediumBad) THEN
        _bSafeLatch := FALSE;                      (* 作用域②：安全恢复才清 E3 / Clear E3 only if safe *)
    END_IF
    _eCause := E_DL_QtlCause.eNone;                (* 作用域③：清成因与分级 / Clear cause and grade *)
    _eGrade := E_DL_QtlGrade.eG0;
    _nRetry := 0;                                  (* 作用域④：清重试 / Clear retry *)
    _fCycleAccS := 0.0;                            (* 作用域⑤：清本件节拍累加 / Clear cycle accumulator *)
    IF NOT _bSafeLatch THEN
        IF (_ePhase = E_DL_QtlPhase.eFault) OR (_ePhase = E_DL_QtlPhase.eSafeStop) THEN
            _ePhase := E_DL_QtlPhase.eIdle;        (* 作用域⑥：故障相迁回待机 / Back to idle *)
        END_IF
    END_IF
ELSIF bStop AND (_ePhase <> E_DL_QtlPhase.eIdle) AND (_ePhase <> E_DL_QtlPhase.eSafeStop) THEN
    IF _ePhase = E_DL_QtlPhase.eFault THEN
        _bFault := FALSE;                          (* 中止清 E2（E3 只能由复位清） / Abort clears E2 only *)
        _eCause := E_DL_QtlCause.eNone;
        _eGrade := E_DL_QtlGrade.eG0;
    END_IF
    _nRetry := 0;                                  (* 重试复位 / Retry reset *)
    _fCycleAccS := 0.0;                            (* 节拍累加作废 / Cycle accumulator void *)
    _ePhase := E_DL_QtlPhase.eIdle;                (* 回待机 / Back to idle *)
END_IF

(* —— 段 5：本件节拍累加（仅工作相计时，故障与安全相不累） —— *)
IF (_ePhase <> E_DL_QtlPhase.eIdle) AND (_ePhase <> E_DL_QtlPhase.eFault) AND (_ePhase <> E_DL_QtlPhase.eSafeStop) THEN
    _fCycleAccS := _fCycleAccS + _fCy;
END_IF

(* —— 段 6：故障请求统一落地（分支内只写成因与请求，落地仅此一处，R187/R252） —— *)
IF _bFaultReq AND (NOT _bSafeLatch) THEN
    _bFault := TRUE;                               (* E2 锁存 / Latch E2 *)
    _eGrade := E_DL_QtlGrade.eG2;                  (* 分级 E2 / Grade E2 *)
    _ePhase := E_DL_QtlPhase.eFault;               (* 同步迁相（R252） / Migrate *)
    bError := TRUE;                                (* 故障标志同段置位（R45 配对） / Error pairing *)
END_IF

(* —— 段 7：主状态机（ENUM + CASE，ELSE 兜底回安全相） —— *)
CASE _ePhase OF
E_DL_QtlPhase.eIdle:
    IF rtStart.Q AND (NOT _bFault) AND (NOT _bSafeLatch) THEN
        _fCycleAccS := 0.0;                        (* 新件起算 / New piece *)
        _ePhase := E_DL_QtlPhase.eLoad;            (* 入上料相 / To loading *)
    END_IF
E_DL_QtlPhase.eLoad:
    IF bPartLoaded THEN
        _ePhase := E_DL_QtlPhase.eHeat;            (* 上料到位 -> 加热 / Loaded, heat *)
    ELSIF tonLoad.Q THEN
        _eCause := E_DL_QtlCause.eLoadTmo;         (* 归因：上料超时 / Cause: load timeout *)
        _bFaultReq := TRUE;
    END_IF
E_DL_QtlPhase.eHeat:
    IF _bPartBad THEN
        _eCause := E_DL_QtlCause.eSigBad;          (* 归因：温度信号非有限 / Cause: signal *)
        _bFaultReq := TRUE;
    ELSIF _bSoakBand THEN
        _ePhase := E_DL_QtlPhase.eSoak;            (* 到保温带 -> 保温 / In band, soak *)
    ELSIF tonHeat.Q THEN
        IF _nRetry < nRetryMax THEN
            _nRetry := _nRetry + 1;                (* E1：可重试，计时器自复位后重计时 / E1 retry *)
            _eGrade := E_DL_QtlGrade.eG1;
            _eCause := E_DL_QtlCause.eHeatTmo;
        ELSE
            _eCause := E_DL_QtlCause.eRetryOver;   (* 归因：重试耗尽 / Cause: retry exhausted *)
            _bFaultReq := TRUE;
        END_IF
    END_IF
E_DL_QtlPhase.eSoak:
    IF tonSoak.Q AND _bSoakBand THEN
        _ePhase := E_DL_QtlPhase.eQuench;          (* 到时且带内 -> 淬火 / Timed and in band, quench *)
    ELSIF tonSoak.Q THEN
        _eCause := E_DL_QtlCause.eSoakTmo;         (* 归因：到时仍带外 / Cause: out of band at timeout *)
        _bFaultReq := TRUE;
    END_IF
E_DL_QtlPhase.eQuench:
    IF tonQuench.Q AND bQuenchImmersion THEN
        _ePhase := E_DL_QtlPhase.eDrain;           (* 浸没到位且到时 -> 沥液 / Immersed and timed *)
    ELSIF tonQuench.Q THEN
        _eCause := E_DL_QtlCause.eQuenchTmo;       (* 归因：到时未浸没 / Cause: not immersed *)
        _bFaultReq := TRUE;
    END_IF
E_DL_QtlPhase.eDrain:
    IF bDrained THEN
        _ePhase := E_DL_QtlPhase.eTemper;          (* 回液到位 -> 回火 / Drained, temper *)
    ELSIF tonDrain.Q THEN
        IF _nRetry < nRetryMax THEN
            _nRetry := _nRetry + 1;                (* E1：可重试 / E1 retry *)
            _eGrade := E_DL_QtlGrade.eG1;
            _eCause := E_DL_QtlCause.eDrainTmo;
        ELSE
            _eCause := E_DL_QtlCause.eRetryOver;   (* 归因：重试耗尽 / Cause: retry exhausted *)
            _bFaultReq := TRUE;
        END_IF
    END_IF
E_DL_QtlPhase.eTemper:
    IF _bTemperBand AND tonTemper.Q THEN
        _ePhase := E_DL_QtlPhase.eCool;            (* 带内且总窗到 -> 冷却 / In band and window done *)
    ELSIF tonTemper.Q THEN
        _eCause := E_DL_QtlCause.eTemperTmo;       (* 归因：回火超时（带内未达） / Cause: temper timeout *)
        _bFaultReq := TRUE;
    END_IF
E_DL_QtlPhase.eCool:
    IF _bPartBad THEN
        _eCause := E_DL_QtlCause.eSigBad;          (* 归因：温度信号非有限 / Cause: signal *)
        _bFaultReq := TRUE;
    ELSIF fPartTempC <= fCoolSetC THEN
        _ePhase := E_DL_QtlPhase.eUnload;          (* 冷到出料温度 -> 下料 / Cooled, unload *)
    ELSIF tonCool.Q THEN
        _eCause := E_DL_QtlCause.eCoolTmo;         (* 归因：冷却超时 / Cause: cool timeout *)
        _bFaultReq := TRUE;
    END_IF
E_DL_QtlPhase.eUnload:
    IF bUnloadPermit THEN
        _bDonePulse := TRUE;                       (* 单拍完成（段 1 预清） / One-scan done *)
        _tCycleLast := CalcCycleTime();            (* 委托方法换算节拍 / Delegate cycle conversion *)
        _fCycleSumS := _fCycleSumS + _fCycleAccS;  (* 节拍总和累加 / Cycle sum *)
        _fCycleAccS := 0.0;                        (* 本件累加清零 / Clear accumulator *)
        IF _nPiece < DL_QTL_PCMAX THEN
            _nPiece := _nPiece + 1;                (* 产量推进（容量载体判上限） / Saturating count *)
        END_IF
        _ePhase := E_DL_QtlPhase.eIdle;            (* 回待机迎下一件 / Back to idle *)
    ELSIF tonUnload.Q THEN
        _eCause := E_DL_QtlCause.eUnloadTmo;       (* 归因：下料超时 / Cause: unload timeout *)
        _bFaultReq := TRUE;
    END_IF
E_DL_QtlPhase.eFault:
    bError := TRUE;                                (* 故障相驻留（锁存回放） / Fault residency *)
E_DL_QtlPhase.eSafeStop:
    bError := TRUE;                                (* 安全相驻留（锁存回放） / Safety residency *)
ELSE
    _eCause := E_DL_QtlCause.ePhaseBad;            (* 非法相位兜底 / Illegal phase fallback *)
    _bFault := TRUE;                               (* 兜底锁存 / Fallback latch *)
    _eGrade := E_DL_QtlGrade.eG2;                  (* 兜底分级 E2 / Fallback grade *)
    _ePhase := E_DL_QtlPhase.eFault;               (* 回安全侧 / Fall back to fault *)
    bError := TRUE;
END_CASE

(* —— 段 8：统一出口（电平量由 _ePhase 派生，单拍量由 _b* 标志映射） —— *)
eState := _ePhase;                                 (* 相出口 / Phase outlet *)
eCause := _eCause;                                 (* 成因回放 / Cause playback *)
eGrade := _eGrade;                                 (* 分级出口 / Grade outlet *)
bError := bError OR _bFault OR _bSafeLatch;        (* 故障标志汇总（E1 不置） / Error summary *)
bSafeCut := _bSafeLatch;                           (* 安全断能指令 / Safety energy cut *)
bHeatActive := (_ePhase = E_DL_QtlPhase.eHeat);    (* 加热相指示 / Heating indicator *)
bQuenchActive := (_ePhase = E_DL_QtlPhase.eQuench);(* 淬火相指示 / Quench indicator *)
bDone := _bDonePulse;                              (* 单拍完成脉冲 / One-scan done *)
nPieceCount := _nPiece;                            (* 产量出口 / Count outlet *)
tCycleLast := _tCycleLast;                         (* 节拍出口 [ms] / Cycle outlet *)
IF _nPiece > 0 THEN
    fCycleAvgS := _fCycleSumS / UDINT_TO_LREAL(_nPiece);   (* 均值分母已判非零 / Guarded mean *)
ELSE
    fCycleAvgS := 0.0;                             (* 无件输出 0 / No piece, zero *)
END_IF
nRetryUsed := _nRetry;                             (* 重试占用出口 / Retry outlet *)
_ePhasePrev := _ePhase;                            (* 段末相快照（下拍迁移后置用） / Phase snapshot *)
END_FUNCTION_BLOCK

(* ---- FB_DL_RadiatorZoneValve.st ---- *)
(*
  FB_DL_RadiatorZoneValve  —  散热器末端温控阀脉冲控制 / Radiator zone valve pulse control
  分类 Category : DL_Process
  码位 Code     : 16#06_0_B9
  段位说明      : R38 W7 预留 B6~BF 本轮正式启用，B8 格由 CartonDenestPush 启用，本件启用 B9 格
  版本 Version  : 1.0.0
  来源 Source   : t2-2-lbp — FB_DL_ThreePointValve 典型消费场景待挖项
  溯源 Origin   : clean-room 实现，三点浮阀 + 房间温度闭环为公开经典控制语义，未复制任何源码行
  功能 Function : 1) 房间温度闭环：FC_DL_Hysteresis 迟滞判热需求（fRoomSpC 设定 + fBandC 回差带，
                  带内保持，防阀频繁切换）；
                  2) FB_DL_ThreePointValve 实例消费：热需求 → 开阀指令，无需求 → 关阀指令；
                  3) 最小启停间隔保护：全开后 tMinRun 内禁关、全关后 tMinOff 内禁开
                  （tonMinRun/tonMinOff 双实例，被闭锁期间置信息级码）；
                  4) 阀门限位开关与行程时间由组态透传，估算开度镜像出口。
  边界 Boundary : ① 本件只出三点阀开关指令（经 FB_DL_ThreePointValve 输出脉冲），不写物理 IO；
                  ② 温度信号非有限：需求冻结保持（不误开不误关）+ 信息级码；
                  ③ R228-A 达标声明：tonMinRun/tonMinOff 各自单用途计时（IN 为单相等式），
                  无跨相复用问题（本件无状态机相）；
                  ④ 组态域闸覆盖全部参与换算引脚（R151）；迟滞带/间隔域非法判组态错锁存；
                  ⑤ 需求判据取反口径：迟滞件 TRUE = 温度高（停热），需求 = NOT 迟滞输出，
                  上电冷态需求为 TRUE（保守供热侧）。
  依赖 Depends  : FB_DL_ThreePointValve（实例化，引脚按 registry 实名）；
                  FC_DL_Hysteresis（函数调用，bState 由本件成员持有回传）
  码表 Error codes（本件格 06_0_B9，子码步进 +0x100）:
    16#0006_01B9 信息级：最小启停间隔闭锁中（指令暂缓，不置故障）
    16#0006_02B9 故障级：组态非法（设定/回差/间隔域非法），锁存至复位
    16#0006_03B9 信息级：温度信号非有限，需求冻结保持
    16#0006_04B9 信息级：加热需求置位（bHeating 拍）
    16#0006_05B9 故障级：保留码，本件无 CASE 主状态机，仅作后续维护者新增分支时的防御式默认码

  修订历史 Revision :
    2026-11-19  v1.0.0  R39 首版（批次 4 · 序号 17）
*)

FUNCTION_BLOCK FB_DL_RadiatorZoneValve
VAR_INPUT
    bEnable      : BOOL := TRUE;       // 总使能，FALSE 时关阀指令并冻结需求 [-] / Master enable
    fRoomTempC   : REAL := 20.0;       // 房间实测温度 [°C] / Room measured temperature
    fRoomSpC     : REAL := 21.0;       // 房间设定温度 [°C] / Room setpoint
    fBandC       : REAL := 0.5;        // 需求回差带 [°C]，域 > 0 / Demand hysteresis band
    bLimOpen     : BOOL := FALSE;      // 阀全开限位反馈（透传三点阀）[-] / Valve open limit, passed through
    bLimClosed   : BOOL := FALSE;      // 阀全关限位反馈（透传三点阀）[-] / Valve closed limit, passed through
    tStrokeOpen  : TIME := T#60S;      // 全行程开启时间 [ms]（透传三点阀）/ Full-open stroke time
    tStrokeClose : TIME := T#60S;      // 全行程关闭时间 [ms]（透传三点阀）/ Full-close stroke time
    tMinRun      : TIME := T#120S;     // 最小运行间隔（全开后禁关时长）[ms]，域 >= 0 / Minimum run time
    tMinOff      : TIME := T#120S;     // 最小停歇间隔（全关后禁开时长）[ms]，域 >= 0 / Minimum off time
    bReset       : BOOL := FALSE;      // 故障复位，上升沿生效 / Fault reset, rising edge
END_VAR
VAR_OUTPUT
    bHeating     : BOOL;               // 加热需求（迟滞后，电平）[-] / Heating demand, level
    bOpenCmd     : BOOL;               // 开阀指令生效中（透传阀件脉冲前）[-] / Open command active
    bCloseCmd    : BOOL;               // 关阀指令生效中 [-] / Close command active
    bOpened      : BOOL;               // 阀全开确认（限位优先）[-] / Valve fully opened
    bClosed      : BOOL;               // 阀全关确认（限位优先）[-] / Valve fully closed
    fValvePosEst : REAL;               // 阀估算开度 [%]（三点阀积分口径）/ Valve estimated position
    bError       : BOOL;               // 故障锁存，仅故障级码置位，bReset 清除 [-] / Fault latch
    uErrorId     : UDINT;              // 事件码，0 = 无事件（故障级锁存回放）/ Event code
END_VAR
VAR
    fbValve    : FB_DL_ThreePointValve;   // 三点浮阀实例（主体首部无条件刷新）/ Three-point valve instance
    tonMinRun  : TON;                     // 最小运行计时（全开期间，单用途）/ Minimum run timer, single purpose
    tonMinOff  : TON;                     // 最小停歇计时（全关期间，单用途）/ Minimum off timer, single purpose
    rtReset    : R_TRIG;                  // 复位上升沿 / Reset rising edge
    _bTempHigh : BOOL;                    // 迟滞判温高回传保持变量 / Hysteresis temp-high hold member
    _bHeatDem  : BOOL := TRUE;            // 热需求内部量（上电冷态为 TRUE，保守供热）/ Internal heat demand, TRUE on cold start
    _bTempBad  : BOOL;                    // 温度非有限标志 / Temperature non-finite flag
    _bOpenReq  : BOOL;                    // 开阀请求（需求 + 间隔闭锁裁决后）/ Open request after gating
    _bCloseReq : BOOL;                    // 关阀请求（需求取反 + 间隔闭锁裁决后）/ Close request after gating
    _bBlocked  : BOOL;                    // 本拍指令被间隔闭锁标志 / Command blocked by interval this cycle
    _bOpenedPrv: BOOL;                    // 上拍全开确认镜像（间隔计时基准）/ Previous fully-open mirror, timer basis
    _bClosedPrv: BOOL;                    // 上拍全关确认镜像（间隔计时基准）/ Previous fully-closed mirror, timer basis
    _uInfo     : UDINT;                   // 信息码，每拍重算 / Info code
    _uFault    : UDINT;                   // 故障码锁存寄存 / Latched fault code register
    _bFault    : BOOL;                    // 故障锁存位 / Latched fault bit
    _bCfgBad   : BOOL;                    // 组态非法聚合 / Configuration invalid aggregate
END_VAR
VAR CONSTANT
    DL_RZV_INF_CAP : REAL := 1.0E15;  // 非有限值筛查幅值上限 / Non-finite screening cap
END_VAR

(* —— 段 0：定时器与边沿实例无条件周期刷新（R182：调用语句不得置于 IF/CASE 内） —— *)
(* 间隔计时 IN 取上拍阀位确认镜像（SemaMutex 同款「IN 取上一拍锁存状态」口径） *)
rtReset(CLK := bReset);                                 // 复位沿刷新，每拍必调
tonMinRun(IN := _bOpenedPrv, PT := tMinRun);            // 最小运行计时（上拍全开电平，单用途）
tonMinOff(IN := _bClosedPrv, PT := tMinOff);            // 最小停歇计时（上拍全关电平，单用途）

(* —— 段 1：单拍量预清零（锁存量 _uFault/_bFault/_bHeatDem/_bTempHigh 不入清单，R187①） —— *)
_uInfo := 16#0000_0000;             // 信息码每拍重算
_bCfgBad := FALSE;                  // 组态非法预清零
_bBlocked := FALSE;                 // 闭锁标志预清零
uErrorId := 16#0000_0000;           // 事件码缺省无事件

(* —— 段 3：组态域闸（覆盖全部参与判据换算的引脚，R151） —— *)
IF (fRoomTempC <> fRoomTempC) OR (ABS(fRoomTempC) > DL_RZV_INF_CAP) OR ((fRoomTempC - fRoomTempC) <> 0.0)
   OR (fRoomSpC <> fRoomSpC) OR (ABS(fRoomSpC) > DL_RZV_INF_CAP) THEN
    _bTempBad := TRUE;              // 温度/设定非有限（需求冻结保持，信息级）
END_IF
IF (fBandC <= 0.0) OR (TIME_TO_DINT(tMinRun) < 0) OR (TIME_TO_DINT(tMinOff) < 0)
   OR (TIME_TO_DINT(tStrokeOpen) <= 0) OR (TIME_TO_DINT(tStrokeClose) <= 0) THEN
    _bCfgBad := TRUE;               // 回差/间隔/行程域非法
END_IF
IF _bCfgBad AND (NOT _bFault) THEN
    _uFault := 16#0006_02B9;        // 故障级：组态非法（仅首次进入时写入）
    _bFault := TRUE;
END_IF
IF rtReset.Q AND (NOT _bCfgBad) THEN
    _bFault := FALSE;               // 清故障锁存位（R228-B：rtReset.Q 恒可达）
    _uFault := 16#0000_0000;
END_IF

(* —— 段 4：需求判定（迟滞取反口径；非有限冻结保持） —— *)
IF (NOT _bTempBad) AND (NOT _bCfgBad) THEN
    _bTempHigh := FC_DL_Hysteresis(fIn := fRoomTempC,       // 迟滞判温高（TRUE = 停热侧）
                                   fThreshold := fRoomSpC,  // 设定点
                                   fHysteresis := fBandC,   // 回差带
                                   bState := _bTempHigh);   // 回传保持变量（同一成员，有状态纪律）
    _bHeatDem := NOT _bTempHigh;    // 需求 = NOT 温高（带内保持，防阀频切）
    IF _bHeatDem THEN
        _uInfo := 16#0006_01B9;     // 信息级：加热需求置位
    END_IF
ELSE
    _uInfo := 16#0006_03B9;         // 信息级：温度信号非有限，需求冻结保持（_bHeatDem 不改写）
END_IF

(* —— 段 5：最小启停间隔裁决（先于三点阀调用，数据流「先算后喂」） —— *)
IF NOT bEnable THEN
    _bOpenReq := FALSE;             // 失能：禁开
    _bCloseReq := TRUE;             // 失能：关阀（安全供热侧）
    _bHeatDem := FALSE;             // 失能：需求清零（出口同步）
ELSIF _bFault THEN
    _bOpenReq := FALSE;             // 故障：禁开
    _bCloseReq := TRUE;             // 故障：关阀（安全侧）
    _bHeatDem := FALSE;             // 故障：需求清零（出口同步）
ELSE
    _bOpenReq := _bHeatDem AND (NOT tonMinOff.Q);   // 开阀 = 需求 AND 非停歇闭锁
    _bCloseReq := (NOT _bHeatDem) AND (NOT tonMinRun.Q);    // 关阀 = 无需求 AND 非运行闭锁
    IF _bHeatDem AND tonMinOff.Q THEN
        _bBlocked := TRUE;          // 开阀被停歇闭锁
    END_IF
    IF (NOT _bHeatDem) AND tonMinRun.Q THEN
        _bBlocked := TRUE;          // 关阀被运行闭锁
    END_IF
END_IF
IF _bBlocked THEN
    _uInfo := 16#0006_01B9;         // 信息级：间隔闭锁中（覆盖需求码，闭锁状态优先）
END_IF

(* —— 段 6：三点阀实例调用（每拍顶层无条件；裁决结果作引脚） —— *)
fbValve(bCmdOpen := _bOpenReq,      // 开阀指令（电平）
        bCmdClose := _bCloseReq,    // 关阀指令（电平；与开同拍为假，裁决互斥）
        bLimOpen := bLimOpen,       // 限位透传
        bLimClosed := bLimClosed,   // 限位透传
        tStrokeOpen := tStrokeOpen, // 行程透传
        tStrokeClose := tStrokeClose,   // 行程透传
        fEstimateTol := 10.0,       // 估算-限位一致性容差（默认口径）
        bEnable := TRUE,            // 阀件动作联锁恒放行（闭锁已在本件裁决）
        bReset := bReset,           // 复位透传
        bTrack := FALSE);           // 不跟踪（限位开关口径由透传承载）

(* —— 段 7：出口单点映射（名实同源；锁存码回放，禁同拍抹除） —— *)
_bOpenedPrv := fbValve.bOpened;     // 上拍全开镜像更新（下一拍间隔计时基准）
_bClosedPrv := fbValve.bClosed;     // 上拍全关镜像更新
bHeating := _bHeatDem;              // 需求出口镜像
bOpenCmd := fbValve.bOpenPulse;     // 开阀脉冲镜像（阀件输出）
bCloseCmd := fbValve.bClosePulse;   // 关阀脉冲镜像
bOpened := fbValve.bOpened;         // 全开确认镜像
bClosed := fbValve.bClosed;         // 全关确认镜像
fValvePosEst := fbValve.fPosEstimate;   // 估算开度镜像
IF _bFault THEN
    uErrorId := _uFault;            // 故障锁存码回放
    bError := TRUE;
ELSE
    uErrorId := _uInfo;             // 信息码
    bError := FALSE;
END_IF

END_FUNCTION_BLOCK

(* ---- FB_DL_ReactorChargeSeq.st ---- *)
(*
  DL Factory R84 | FB_DL_ReactorChargeSeq
  功能：反应釜多组分投料顺序时序，逐相流量累积达标判据与搅拌运行互锁
  开源溯源：无（clean-room 自研，依据公开工艺公式，来源=行业通用公式，许可证=MIT，借鉴点=公式结构）
  规则：R1-R16 全遵守
*)
TYPE E_DL_RctChgState :
(
    eIdle := 0, // 空闲待启动 [-] / idle [-]
    eStirCheck := 1, // 搅拌运行确认相 [-] / stirrer check phase [-]
    eChargeA := 2, // A 组分投料相 [-] / component A charging phase [-]
    eChargeB := 3, // B 组分投料相 [-] / component B charging phase [-]
    eChargeC := 4, // C 组分投料相 [-] / component C charging phase [-]
    eHold := 5, // 投料后保持相 [-] / post charge hold phase [-]
    eDone := 6, // 完成相 [-] / done phase [-]
    eFault := 7 // 故障锁存相 [-] / fault latched phase [-]
) := eIdle;
END_TYPE

FUNCTION_BLOCK FB_DL_ReactorChargeSeq
VAR_INPUT
    xStart : BOOL; // 投料启动按钮 [-] / charge start pushbutton [-]
    xReset : BOOL; // 复位按钮，上升沿清故障码与累积量 [-] / reset pushbutton [-]
    xStirRunning : BOOL; // 搅拌运行反馈（投料互锁条件） [-] / stirrer running interlock feedback [-]
    fFlowKgh : REAL; // 当前投料瞬时流量 [kg/h] / instantaneous charge flow [kg/h]
    tScan : TIME := T#50MS; // 扫描周期（累积用） [s] / scan period for accumulation [s]
    aTargetKg : ARRAY[0..2] OF REAL; // A/B/C 三组分目标投料量 [kg] / target mass per component [kg]
    tStirLimit : TIME := T#10S; // 搅拌确认超时 [s] / stirrer check timeout [s]
    tPhaseLimit : TIME := T#600S; // 单组分投料相超时 [s] / per component charge timeout [s]
    tHoldLimit : TIME := T#120S; // 投料后保持时长 [s] / post charge hold duration [s]
END_VAR
VAR_OUTPUT
    eState : E_DL_RctChgState; // 当前时序状态 [-] / current sequence state [-]
    iErrCode : INT; // 故障码 0=正常，501~506 [-] / error code, 501 to 506 [code]
    fChargedKg : REAL; // 本批已投料累计质量 [kg] / total charged mass of this batch [kg]
    xDone : BOOL; // 完成单拍脉冲 [-] / done one-shot pulse [-]
END_VAR
VAR
    rtStart : R_TRIG; // 启动上升沿实例 [-] / start rising edge instance [-]
    rtReset : R_TRIG; // 复位上升沿实例 [-] / reset edge instance [-]
    tonStir : TON; // 搅拌确认超时定时器 [-] / stirrer check timer [-]
    tonPhaseA : TON; // A 组分投料超时定时器（各相独立，R571） [-] / component A charge timer, one per phase [-]
    tonPhaseB : TON; // B 组分投料超时定时器（各相独立，R571） [-] / component B charge timer, one per phase [-]
    tonPhaseC : TON; // C 组分投料超时定时器（各相独立，R571） [-] / component C charge timer, one per phase [-]
    tonHold : TON; // 保持相定时器 [-] / hold phase timer [-]
    _eState : E_DL_RctChgState := E_DL_RctChgState.eIdle; // 内部相位（CASE 唯一写目标） [-] / internal phase [-]
    _iErr : INT; // 故障码内部锁存 [-] / latched error code [-]
    fCharged : REAL; // 累计投料量内部量 [kg] / internal charged mass [kg]
    fPhaseKg : REAL; // 当前组分已投量 [kg] / mass charged in the current phase [kg]
    fDtSec : REAL; // 扫描周期秒值 [s] / scan period in seconds [s]
    fStepKg : REAL; // 本拍投料增量 [kg] / charge increment of this scan [kg]
    xDoneInt : BOOL; // 完成内部锁存位 [-] / internal done latch [-]
    xDonePrev : BOOL; // 完成前拍快照 [-] / done previous scan snapshot [-]
END_VAR

// 段 0｜边沿与定时器实例无条件周期刷新（R7）
rtStart(CLK := xStart); // 启动沿每拍必调 [-] / start edge every scan [-]
rtReset(CLK := xReset); // 复位沿每拍必调 [-] / reset edge every scan [-]
tonStir(IN := _eState = E_DL_RctChgState.eStirCheck, PT := tStirLimit); // 搅拌确认相闸 [-] / stirrer check phase gate [-]
tonPhaseA(IN := _eState = E_DL_RctChgState.eChargeA, PT := tPhaseLimit); // A 相独立计时，离相即复位 [-] / component A timer, reset when the phase leaves [-]
tonPhaseB(IN := _eState = E_DL_RctChgState.eChargeB, PT := tPhaseLimit); // B 相独立计时，离相即复位 [-] / component B timer, reset when the phase leaves [-]
tonPhaseC(IN := _eState = E_DL_RctChgState.eChargeC, PT := tPhaseLimit); // C 相独立计时，离相即复位 [-] / component C timer, reset when the phase leaves [-]
tonHold(IN := _eState = E_DL_RctChgState.eHold, PT := tHoldLimit); // 保持相闸 [-] / hold phase gate [-]

// 段 1｜本拍增量派生（kg/h × s ÷ 3600 = kg）
fDtSec := LREAL_TO_REAL(TIME_TO_LREAL(tScan) / 1000.0); // ms ÷ 1000 = s / [ms] / 1000 = [s]
fStepKg := 0.0; // 增量初值零 [kg] / increment starts at zero [kg]
IF (fFlowKgh > -1.0E30 AND fFlowKgh < 1.0E30) AND fFlowKgh > 0.0 THEN
    fStepKg := (fFlowKgh * fDtSec) / 3600.0; // kg/h × s ÷ 3600 s/h = kg / [kg/h] × [s] / 3600 = [kg]
END_IF

// 段 2｜复位沿：清故障码、累积量与相位（R189）
IF rtReset.Q THEN
    _iErr := 0; // 清故障码 [-] / clear error code [-]
    fCharged := 0.0; // 清本批累计投料 [kg] / clear the batch charge [kg]
    fPhaseKg := 0.0; // 清当前组分累计 [kg] / clear the phase charge [kg]
    xDoneInt := FALSE; // 清完成锁存 [-] / clear done latch [-]
    _eState := E_DL_RctChgState.eIdle; // 回空闲相 [-] / back to idle [-]
END_IF

// 段 3｜主状态机（合法事件优先于超时迁移，R275）
CASE _eState OF
    E_DL_RctChgState.eIdle: // 空闲相 [-] / idle [-]
        xDoneInt := FALSE; // 空闲清完成锁存 [-] / clear done latch in idle [-]
        fCharged := 0.0; // 空闲期累计归零 [kg] / hold the accumulator at zero [kg]
        fPhaseKg := 0.0; // 空闲期组分累计归零 [kg] / hold the phase accumulator at zero [kg]
        IF rtStart.Q THEN
            _eState := E_DL_RctChgState.eStirCheck; // 启动沿先确认搅拌 [-] / start edge checks the stirrer [-]
        END_IF
    E_DL_RctChgState.eStirCheck: // 搅拌确认相（互锁：未运行禁投料） [-] / stirrer check [-]
        IF xStirRunning AND NOT tonStir.Q THEN
            _eState := E_DL_RctChgState.eChargeA; // 搅拌运行转 A 组分 [-] / stirrer running leads to component A [-]
        ELSIF tonStir.Q THEN
            _iErr := 501; _eState := E_DL_RctChgState.eFault; // 搅拌未运行超时（禁投料） [-] / stirrer timeout, charging blocked [-]
        END_IF
    E_DL_RctChgState.eChargeA: // A 组分投料相 [-] / component A [-]
        IF NOT xStirRunning THEN
            _iErr := 502; _eState := E_DL_RctChgState.eFault; // 投料中搅拌停转（互锁断开） [-] / stirrer lost during charging [-]
        ELSIF fPhaseKg >= aTargetKg[0] THEN
            fPhaseKg := 0.0; // 本组分累计清零 [kg] / clear the phase accumulator [kg]
            _eState := E_DL_RctChgState.eChargeB; // A 达标转 B [-] / A reached leads to B [-]
        ELSIF tonPhaseA.Q THEN
            _iErr := 503; _eState := E_DL_RctChgState.eFault; // A 组分投料超时 [-] / component A timeout [-]
        ELSE
            fCharged := fCharged + fStepKg; // kg + kg = kg / [kg] + [kg] = [kg]
            fPhaseKg := fPhaseKg + fStepKg; // kg + kg = kg / [kg] + [kg] = [kg]
        END_IF
    E_DL_RctChgState.eChargeB: // B 组分投料相 [-] / component B [-]
        IF NOT xStirRunning THEN
            _iErr := 502; _eState := E_DL_RctChgState.eFault; // 投料中搅拌停转 [-] / stirrer lost during charging [-]
        ELSIF fPhaseKg >= aTargetKg[1] THEN
            fPhaseKg := 0.0; // 本组分累计清零 [kg] / clear the phase accumulator [kg]
            _eState := E_DL_RctChgState.eChargeC; // B 达标转 C [-] / B reached leads to C [-]
        ELSIF tonPhaseB.Q THEN
            _iErr := 504; _eState := E_DL_RctChgState.eFault; // B 组分投料超时 [-] / component B timeout [-]
        ELSE
            fCharged := fCharged + fStepKg; // kg + kg = kg / [kg] + [kg] = [kg]
            fPhaseKg := fPhaseKg + fStepKg; // kg + kg = kg / [kg] + [kg] = [kg]
        END_IF
    E_DL_RctChgState.eChargeC: // C 组分投料相 [-] / component C [-]
        IF NOT xStirRunning THEN
            _iErr := 502; _eState := E_DL_RctChgState.eFault; // 投料中搅拌停转 [-] / stirrer lost during charging [-]
        ELSIF fPhaseKg >= aTargetKg[2] THEN
            fPhaseKg := 0.0; // 本组分累计清零 [kg] / clear the phase accumulator [kg]
            _eState := E_DL_RctChgState.eHold; // C 达标转保持相 [-] / C reached leads to hold [-]
        ELSIF tonPhaseC.Q THEN
            _iErr := 505; _eState := E_DL_RctChgState.eFault; // C 组分投料超时 [-] / component C timeout [-]
        ELSE
            fCharged := fCharged + fStepKg; // kg + kg = kg / [kg] + [kg] = [kg]
            fPhaseKg := fPhaseKg + fStepKg; // kg + kg = kg / [kg] + [kg] = [kg]
        END_IF
    E_DL_RctChgState.eHold: // 保持相：搅拌必须仍在运行 [-] / hold phase [-]
        IF NOT xStirRunning THEN
            _iErr := 502; _eState := E_DL_RctChgState.eFault; // 保持期搅拌停转 [-] / stirrer lost during hold [-]
        ELSIF tonHold.Q THEN
            _eState := E_DL_RctChgState.eDone; // 保持时长到转完成相 [-] / hold done leads to done [-]
        END_IF
    E_DL_RctChgState.eDone: // 完成相 [-] / done [-]
        xDoneInt := TRUE; // 置完成锁存（出口统一映射单拍） [-] / raise done latch [-]
        IF NOT xStart THEN
            _eState := E_DL_RctChgState.eIdle; // 松开启动即回空闲 [-] / start released returns to idle [-]
        END_IF
    E_DL_RctChgState.eFault: // 故障相：码值锁存回放，仅复位沿出 [-] / fault, exit only on reset [-]
        ; // 锁存回放（R28） [-] / replay the latch only [-]
ELSE
    _iErr := 506; _eState := E_DL_RctChgState.eFault; // 非法相位兜底 [-] / illegal phase fallback [-]
END_CASE

// 段 4｜出口映射（名实双出口，同源赋值）
eState := _eState; // 状态出口 [-] / state outlet [-]
iErrCode := _iErr; // 故障码出口（锁存值） [-] / error code outlet [-]
fChargedKg := fCharged; // 累计投料出口 [kg] / charged mass outlet [kg]
xDone := xDoneInt AND NOT xDonePrev; // 完成单拍（内部锁存 → 出口映射） [-] / done one-shot [-]
xDonePrev := xDoneInt; // 本拍快照供下拍比较 [-] / snapshot for the next scan [-]
END_FUNCTION_BLOCK

(* ---- FB_DL_ReactorRunawayGuard.st ---- *)
(*
  DL Factory R84 | FB_DL_ReactorRunawayGuard
  功能：间歇反应釜放热失控五级联锁：温升速率、绝热温升外推 MTSR、冷却能力失效三判据并行分档，合成 0~5 级动作需求；升级立即生效、降级按延时逐级回落，五级动作位互斥且可降级；L5 全停锁存至复位沿。
  开源溯源：无（clean-room 自研，依据公开工艺公式与安全设计惯例，来源=行业通用公式+工程实践，许可证=MIT，借鉴点=公式结构与联锁分层）
  规则：R1-R16 全遵守
  ------------------------------------------------------------------
  分类 DL_Process ｜ 复杂度 cx5 ｜ 版本 v1.0.0 ｜ 平台 纯 IEC 61131-3（TON、R_TRIG、LREAL、ENUM、CASE）
  边界一：只出分级动作位与诊断量，不驱动泄放阀、冷却阀与投料阀本体，不采集变送器（属主边界，执行由下层 PRG 完成）。
  边界二：三判据分档——判据①温升速率按 fRateTripKmin 的 0.50/0.65/0.80/0.92/1.00 五档；判据②MTSR 按安全裕度 fMtsrMarginK 的已耗比例 0.50/0.35/0.20/0.08/0.00 五档；
          判据③冷却能力按流量下限与夹套-进水温差反向分 3 档与 4 档，温差反向且流量低于半限时直接判 5 档。
  边界三：MTSR 公式＝反应温度 ＋ 累积投料若全部反应的绝热温升：ΔTad [K]＝|ΔH| [kJ/mol] × 1000 [mol/kmol] × 累积摩尔数 [kmol] ÷（批量 [kg] × cp [kJ/(kg·K)]），
          累积摩尔数 [kmol]＝累积投料 [kg] ÷ 平均摩尔质量 [kg/kmol]；ΔTad 上限兜底 300 K 防外推发散。
  边界四：平均摩尔质量 DL_RAG_MOLAR_KGKMOL 为物料体系代理常量——代理值是反应主料的平均摩尔质量、覆盖 100~200 g/mol 的常规精细化工体系、
          体系外（聚合/无机盐）由上层以实测绝热温升标定后换算入参负责（R95 三句齐备，代理假设挂编译验证债）。
  边界五：分级互斥与可降级——iStage 为唯一权威（0~5 整数），五级位按 xStageN＝(iStage ≥ N) 单源派生；升级无延时（安全侧优先），
          降级由 tDegrade 周期窗逐级回落，窗为自复位形式（IN 串 NOT 自身 Q，R188），故不存在同拍双窗，R100 配比约束不适用（本件只有一件定时器）。
  边界六：相位由分级单源映射、零滞后（R191 名实同源），不设独立相位状态机与分级机双权威。
  安全侧：任一浮点入参非有限、组态越域、或任一判据达 5 档 → 立即迁 eTrip 并锁存 xTripLatched；锁存唯一解除路径为 bReset 上升沿（R188），其余路径（失能、条件消失）均不解锁。
  码表：故障级 2711 入参非有限、2712 组态越域、2713 温升速率达 5 档、2714 MTSR 达 5 档、2715 冷却完全失效、2716 非法分级值（防御性保留）；
        以上六码锁存回放且置 bError（R45 配对）；信息级 2701~2705＝当前分级（1~5 级）之动作码，每拍重算且不置 bError。
  输出契约：xStage1..xStage5 为累积电平（N 级生效则 1..N 位全真，互斥性由 iStage 单源保证）；xAlarmOut/xFeedStop/xMaxCool/xVentCmd/xTotalStop 与分级同源派生；
          fMtsrC/fRateKmin/fDtAdK 为诊断连续量，非有限时出零不外抛；xValid 在锁存或闸不过时为假。
  修订记录：2026-11-24 v1.0.0 R84 首版（批 R84 · 序号 42）
*)

TYPE E_DL_RagState :
(
    eNormal   := 0, // 正常：零级，无动作 / normal, level zero, no action
    eWarn     := 1, // 报警：一级，仅告知 / warn, level one, notification only
    eStopFeed := 2, // 停止投料：二级 / stop feeding, level two
    eMaxCool  := 3, // 加大冷却：三级 / maximum cooling, level three
    eVent     := 4, // 紧急泄放：四级 / emergency venting, level four
    eTrip     := 5  // 全停：五级，锁存至复位沿 / total trip, level five, latched until the reset edge
);
END_TYPE

TYPE E_DL_RagCause :
(
    eNone      := 0, // 无成因 / no cause
    eNotFinite := 1, // 入参非有限（故障级 2711）/ a non-finite input, fault grade 2711
    eCfgBad    := 2, // 组态越域（故障级 2712）/ the configuration is out of its domain, fault grade 2712
    eRateHigh  := 3, // 温升速率达五档（故障级 2713）/ the temperature rate reached level five, fault grade 2713
    eMtsrHigh  := 4, // MTSR 达五档（故障级 2714）/ the MTSR reached level five, fault grade 2714
    eCoolLoss  := 5, // 冷却完全失效（故障级 2715）/ the cooling capability was lost, fault grade 2715
    eStageBad  := 6  // 非法分级值（故障级 2716，防御性保留）/ an illegal stage value, fault grade 2716
);
END_TYPE

FUNCTION_BLOCK FB_DL_ReactorRunawayGuard
VAR CONSTANT
    DL_RAG_SEC_MIN     : LREAL := 60.0;    // 秒到分钟折算系数 [s/min] / the second to minute factor [s/min]
    DL_RAG_DT_MIN      : LREAL := 0.001;   // 采样周期下限（速率分母零闸）[s] / the sample period lower bound [s]
    DL_RAG_RATE_ALPHA  : LREAL := 0.30;    // 速率一阶滤波系数 [-] / the first order gain of the rate filter [-]
    DL_RAG_L1_FRAC     : LREAL := 0.50;    // 判据①一级档位系数（跳闸速率的倍数）[-] / the level one factor of the rate criterion [-]
    DL_RAG_L2_FRAC     : LREAL := 0.65;    // 判据①二级档位系数 [-] / the level two factor of the rate criterion [-]
    DL_RAG_L3_FRAC     : LREAL := 0.80;    // 判据①三级档位系数 [-] / the level three factor of the rate criterion [-]
    DL_RAG_L4_FRAC     : LREAL := 0.92;    // 判据①四级档位系数 [-] / the level four factor of the rate criterion [-]
    DL_RAG_M1_FRAC     : LREAL := 0.50;    // 判据②一级档位（裕度已耗比例）[-] / the level one factor of the MTSR criterion [-]
    DL_RAG_M2_FRAC     : LREAL := 0.35;    // 判据②二级档位 [-] / the level two factor of the MTSR criterion [-]
    DL_RAG_M3_FRAC     : LREAL := 0.20;    // 判据②三级档位 [-] / the level three factor of the MTSR criterion [-]
    DL_RAG_M4_FRAC     : LREAL := 0.08;    // 判据②四级档位 [-] / the level four factor of the MTSR criterion [-]
    DL_RAG_COOL_DT_MIN : LREAL := 2.0;     // 夹套与进水温差下限（低于即冷却不足）[K] / the jacket to inlet temperature difference floor [K]
    DL_RAG_FLOW_L4_FRAC: LREAL := 0.50;    // 判据③四级档位流量系数（下限倍数）[-] / the level four flow factor of the cooling criterion [-]
    DL_RAG_DTAD_MAX    : LREAL := 300.0;   // 绝热温升外推上限兜底 [K] / the adiabatic rise extrapolation upper clamp [K]
    DL_RAG_FRAC_MAX    : LREAL := 1.50;    // 已投料占比上限（外推兜底）[-] / the charged fraction upper clamp [-]
    DL_RAG_MOLAR_KGKMOL: LREAL := 100.0;   // 平均摩尔质量代理常量 [kg/kmol] / the mean molar mass proxy [kg/kmol]
    DL_RAG_MOL_PER_KMOL: LREAL := 1000.0;  // 摩尔到千摩尔折算系数 [mol/kmol] / the mole to kilomole factor [mol/kmol]
    DL_RAG_EPS         : LREAL := 1.0E-9;  // 除法零闸与零判定门限 [-] / the division guard and zero test threshold [-]
END_VAR
VAR_INPUT
    bEnable      : BOOL := TRUE;     // 使能，失能只回零级不解除锁存 [-] / enable, a disable only clears the stage and never the latch
    bReset       : BOOL := FALSE;   // 复位上升沿清全停锁存（唯一解除路径）[-] / reset rising edge clears the trip latch, the only release path
    xStirRun     : BOOL := TRUE;    // 搅拌运行反馈，停搅即二级以上 [-] / the agitator running feedback, a stop forces level two or higher
    fTreactC     : LREAL := 25.0;   // 反应温度 [°C] / the reaction temperature [°C]
    fTjacketC    : LREAL := 25.0;   // 夹套温度 [°C] / the jacket temperature [°C]
    fCoolFlowM3h : LREAL := 10.0;   // 冷却水流量 [m³/h] / the cooling water flow [m3/h]
    fCoolInC     : LREAL := 20.0;   // 冷却水进水温度 [°C] / the cooling water inlet temperature [°C]
    fAccumKg     : LREAL := 0.0;    // 累积投料质量（尚未反应部分）[kg] / the accumulated charged mass still unreacted [kg]
    fBatchKg     : LREAL := 1000.0; // 批量总质量 [kg] / the total batch mass [kg]
    fDhKjMol     : LREAL := 80.0;   // 反应焓变（取绝对值参与外推）[kJ/mol] / the reaction enthalpy, the absolute value is used [kJ/mol]
    fCpKjKgK     : LREAL := 3.50;   // 反应液比热容 [kJ/(kg·K)] / the reaction mixture specific heat [kJ/(kg*K)]
    fRateTripKmin: LREAL := 3.00;   // 温升速率跳闸值（五档基准）[K/min] / the rate trip value, the level five base [K/min]
    fMtsrLimitC  : LREAL := 180.0;  // MTSR 安全极限温度 [°C] / the MTSR safety limit temperature [°C]
    fMtsrMarginK : LREAL := 20.0;   // MTSR 安全裕度（分级带宽）[K] / the MTSR safety margin, the staging band [K]
    fFlowMinM3h  : LREAL := 4.00;   // 冷却水流量下限 [m³/h] / the cooling water flow floor [m3/h]
    fDtSec       : LREAL := 0.10;   // 温度采样周期（速率分母）[s] / the temperature sample period, the rate denominator [s]
    tDegrade     : TIME := T#30S;   // 分级降级延时（逐级回落窗）[毫秒] / the stage downgrade delay per step [ms]
END_VAR
VAR_OUTPUT
    eState       : E_DL_RagState := E_DL_RagState.eNormal; // 相位出口（由分级单源映射）[枚举] / the phase outlet mapped from the stage [enum]
    iStage       : INT := 0;      // 当前动作级（0~5，唯一权威）[级] / the active stage, the single authority [level]
    iErrCode     : INT := 0;      // 错误码（故障级锁存回放，信息级每拍重算）[码] / the error code, latched faults and scan info [code]
    bError       : BOOL := FALSE; // 故障标志（与故障级码同源）[-] / the fault flag sharing the fault code source
    xTripLatched : BOOL := FALSE; // 全停锁存（仅复位沿清除）[-] / the trip latch, cleared by the reset edge only
    xValid       : BOOL := FALSE; // 本拍输入与组态可信 [-] / the inputs and the configuration are trustworthy
    xStage1      : BOOL := FALSE; // 一级动作位：报警 [-] / level one action, the alarm
    xStage2      : BOOL := FALSE; // 二级动作位：停止投料 [-] / level two action, stop the feed
    xStage3      : BOOL := FALSE; // 三级动作位：加大冷却 [-] / level three action, maximum cooling
    xStage4      : BOOL := FALSE; // 四级动作位：紧急泄放 [-] / level four action, emergency venting
    xStage5      : BOOL := FALSE; // 五级动作位：全停 [-] / level five action, total trip
    xAlarmOut    : BOOL := FALSE; // 报警输出（一级及以上）[-] / the alarm output from level one on
    xFeedStop    : BOOL := FALSE; // 停止投料输出（二级及以上）[-] / the feed stop output from level two on
    xMaxCool     : BOOL := FALSE; // 加大冷却输出（三级及以上）[-] / the maximum cooling output from level three on
    xVentCmd     : BOOL := FALSE; // 紧急泄放输出（四级及以上）[-] / the emergency vent output from level four on
    xTotalStop   : BOOL := FALSE; // 全停输出（五级）[-] / the total stop output at level five
    fMtsrC       : LREAL := 0.0;  // MTSR 外推值 [°C] / the extrapolated MTSR [°C]
    fRateKmin    : LREAL := 0.0;  // 滤波后温升速率 [K/min] / the filtered temperature rise rate [K/min]
    fDtAdK       : LREAL := 0.0;  // 绝热温升外推量 [K] / the adiabatic rise extrapolation [K]
END_VAR
VAR
    rtReset    : R_TRIG; // 复位沿实例（无量纲）[-] / the reset edge refreshed unconditionally
    tonDown    : TON;    // 降级窗实例（无量纲）[-] / the self resetting downgrade window, its own output inverted
    _eState    : E_DL_RagState := E_DL_RagState.eNormal; // 内部相位（枚举，无量纲）[-] / the internal phase
    _eCause    : E_DL_RagCause := E_DL_RagCause.eNone; // 故障级成因（枚举，无量纲）[-] / the fault cause latched until the reset edge
    _iStage    : INT := 0;  // 内部分级（唯一权威）[级] / the internal stage, the single authority [level]
    _iReq      : INT := 0;  // 三判据合成后的动作需求级 [级] / the aggregated stage demand [level]
    _iNeed     : INT := 0;  // 单判据档位暂存 [级] / the per criterion stage scratch [level]
    _iErrTmp   : INT := 0;  // 本拍码位暂存 [码] / the scan code scratch [code]
    _iErrLch   : INT := 0;  // 故障级码位锁存槽 [码] / the latched fault code [code]
    _bTrip     : BOOL := FALSE; // 全停锁存位 [-] / the trip latch
    _bInit     : BOOL := FALSE; // 首扫初始化完成标志（R310）[-] / the first scan initialisation flag
    _bFinOk    : BOOL := FALSE; // 全部浮点入参有限 [-] / every floating input is finite
    _bCfgOk    : BOOL := FALSE; // 组态参数域内 [-] / the configuration is inside its domain
    _bRateL5   : BOOL := FALSE; // 判据①达五档（独立成因标志，R190）[-] / criterion one reached level five
    _bMtsrL5   : BOOL := FALSE; // 判据②达五档（独立成因标志）[-] / criterion two reached level five
    _bCoolL5   : BOOL := FALSE; // 判据③冷却完全失效（独立成因标志）[-] / criterion three lost the cooling entirely
    _bRateL1   : BOOL := FALSE; // 判据①达一档 [-] / criterion one reached level one
    _bRateL2   : BOOL := FALSE; // 判据①达二档 [-] / criterion one reached level two
    _bRateL3   : BOOL := FALSE; // 判据①达三档 [-] / criterion one reached level three
    _bRateL4   : BOOL := FALSE; // 判据①达四档 [-] / criterion one reached level four
    _fTprev    : LREAL := 0.0;  // 上拍反应温度快照（差分用）[°C] / the previous scan temperature snapshot [°C]
    _fRateRaw  : LREAL := 0.0;  // 原始温升速率（差分值）[K/min] / the raw temperature rise rate [K/min]
    _fRateFilt : LREAL := 0.0;  // 滤波后温升速率（保持槽）[K/min] / the filtered rate, a hold slot [K/min]
    _fFrac     : LREAL := 0.0;  // 累积投料占批量比（钳定后）[-] / the charged fraction after clamping [-]
    _fMoles    : LREAL := 0.0;  // 累积投料摩尔数 [kmol] / the accumulated moles [kmol]
    _fHeatKj   : LREAL := 0.0;  // 累积物料若全部反应放热 [kJ] / the heat if all charged mass reacted [kJ]
    _fDtAd     : LREAL := 0.0;  // 绝热温升外推量（钳定后）[K] / the adiabatic rise after clamping [K]
    _fMtsr     : LREAL := 0.0;  // MTSR 外推温度 [°C] / the extrapolated MTSR [°C]
    _fCoolDt   : LREAL := 0.0;  // 夹套与冷却水进水温差 [K] / the jacket to inlet difference [K]
    _fRateThr1 : LREAL := 0.0;  // 判据①一档门限 [K/min] / the level one rate threshold [K/min]
    _fRateThr2 : LREAL := 0.0;  // 判据①二档门限 [K/min] / the level two rate threshold [K/min]
    _fRateThr3 : LREAL := 0.0;  // 判据①三档门限 [K/min] / the level three rate threshold [K/min]
    _fRateThr4 : LREAL := 0.0;  // 判据①四档门限 [K/min] / the level four rate threshold [K/min]
    _fMtsrThr1 : LREAL := 0.0;  // 判据②一档门限 [°C] / the level one MTSR threshold [°C]
    _fMtsrThr2 : LREAL := 0.0;  // 判据②二档门限 [°C] / the level two MTSR threshold [°C]
    _fMtsrThr3 : LREAL := 0.0;  // 判据②三档门限 [°C] / the level three MTSR threshold [°C]
    _fMtsrThr4 : LREAL := 0.0;  // 判据②四档门限 [°C] / the level four MTSR threshold [°C]
    _tDegrade  : TIME := T#1S;  // 降级窗实参（钳定后）[毫秒] / the downgrade window passed to the timer [ms]
END_VAR
// 段 0｜出口预置：全部出口先赋安全侧值，任何路径不留未初始化输出（安全侧＝全停动作位）/
xValid := FALSE; // 有效性预置假 / validity preset false
xStage1 := FALSE; xStage2 := FALSE; xStage3 := FALSE; // 一至三级位预置假 / levels one to three preset false
xStage4 := FALSE; xStage5 := FALSE; // 四至五级位预置假 / levels four and five preset false
xAlarmOut := FALSE; xFeedStop := FALSE; xMaxCool := FALSE; xVentCmd := FALSE; xTotalStop := FALSE; // 五个动作输出预置假 / the five action outputs preset false
xTripLatched := _bTrip; // 全停锁存回放 / replay the trip latch
iStage := 0; // 分级预置零级，段 11 单点覆盖 / the stage preset zero and overwritten at the outlet
iErrCode := 0; // 码位预置零 / the code preset zero
bError := FALSE; // 故障标志预置假 / the fault flag preset false
fMtsrC := 0.0; fRateKmin := 0.0; fDtAdK := 0.0; // 三个连续量出口预置零 / the three continuous outlets preset zero
eState := E_DL_RagState.eNormal; // 相位预置正常相 / the phase preset normal
_iErrTmp := 0; _iNeed := 0; _iReq := 0; // 单拍暂存预清零（FB32-1：仅单拍变量可预清）/ preclear the scan scratches only
// 段 1｜非有限闸：NaN 自反比较、Inf 差值自减双判，逐项枚举十个浮点入参与两个换算量（R79、R272）
_bFinOk := (fTreactC = fTreactC) AND ((fTreactC - fTreactC) = (fTreactC - fTreactC)) // 反应温度有限 [-] / the reaction temperature is finite
    AND (fTjacketC = fTjacketC) AND ((fTjacketC - fTjacketC) = (fTjacketC - fTjacketC)) // 夹套温度有限 [-] / the jacket temperature is finite
    AND (fCoolFlowM3h = fCoolFlowM3h) AND ((fCoolFlowM3h - fCoolFlowM3h) = (fCoolFlowM3h - fCoolFlowM3h)) // 冷却流量有限 [-] / the cooling flow is finite
    AND (fCoolInC = fCoolInC) AND ((fCoolInC - fCoolInC) = (fCoolInC - fCoolInC)) // 进水温度有限 [-] / the inlet temperature is finite
    AND (fAccumKg = fAccumKg) AND ((fAccumKg - fAccumKg) = (fAccumKg - fAccumKg)) // 累积投料有限 [-] / the accumulated mass is finite
    AND (fBatchKg = fBatchKg) AND ((fBatchKg - fBatchKg) = (fBatchKg - fBatchKg)) // 批量有限 [-] / the batch mass is finite
    AND (fDhKjMol = fDhKjMol) AND ((fDhKjMol - fDhKjMol) = (fDhKjMol - fDhKjMol)) // 焓变有限 [-] / the enthalpy is finite
    AND (fCpKjKgK = fCpKjKgK) AND ((fCpKjKgK - fCpKjKgK) = (fCpKjKgK - fCpKjKgK)) // 比热容有限 [-] / the specific heat is finite
    AND (fRateTripKmin = fRateTripKmin) AND ((fRateTripKmin - fRateTripKmin) = (fRateTripKmin - fRateTripKmin)) // 速率跳闸值有限 [-] / the rate trip value is finite
    AND (fMtsrLimitC = fMtsrLimitC) AND ((fMtsrLimitC - fMtsrLimitC) = (fMtsrLimitC - fMtsrLimitC)) // MTSR 极限有限 [-] / the MTSR limit is finite
    AND (fMtsrMarginK = fMtsrMarginK) AND ((fMtsrMarginK - fMtsrMarginK) = (fMtsrMarginK - fMtsrMarginK)) // 裕度有限 [-] / the margin is finite
    AND (fFlowMinM3h = fFlowMinM3h) AND ((fFlowMinM3h - fFlowMinM3h) = (fFlowMinM3h - fFlowMinM3h)) // 流量下限有限 [-] / the flow floor is finite
    AND (fDtSec = fDtSec) AND ((fDtSec - fDtSec) = (fDtSec - fDtSec)); // 采样周期有限 [-] / the sample period is finite
// 段 2｜组态域闸：全部参与判据换算的限值引脚（R151、FB51-2）
_bCfgOk := (ABS(fRateTripKmin) > DL_RAG_EPS) AND (fMtsrMarginK > DL_RAG_EPS) // 速率跳闸值与裕度非零 [-] / the rate trip and the margin are non zero
    AND (ABS(fFlowMinM3h) > DL_RAG_EPS) AND (fBatchKg > DL_RAG_EPS) // 流量下限与批量非零 [-] / the flow floor and the batch are non zero
    AND (fCpKjKgK > DL_RAG_EPS) AND (fDtSec > DL_RAG_DT_MIN) // 比热容与采样周期域闸 [-] / the specific heat and the sample period gates
    AND (fMtsrLimitC > DL_RAG_EPS) AND (tDegrade > T#0S); // MTSR 极限与降级窗域闸 [-] / the MTSR limit and the window gates
_tDegrade := tDegrade; // 降级窗一级回退：取引脚值 [ms] / level one fallback, take the pin value [ms]
IF _tDegrade <= T#0S THEN _tDegrade := T#1S; END_IF // 降级窗二级回退：按有效域钳定（最小一窗）/ level two, clamp into the valid domain
// 段 3｜首扫初始化与复位沿同块，作用域逐项声明（R310、R311、R152）
IF (NOT _bInit) OR rtReset.Q THEN // 首扫一拍或复位沿 / the first scan or the reset edge
    _bInit := TRUE; // 首扫完成标志（复位沿重复置位同效）/ the first scan flag, the same effect on reset
    _bTrip := FALSE; _eCause := E_DL_RagCause.eNone; _iErrLch := 0; // 作用域一：清全停锁存、清成因、清故障码槽 / scope one, clear the latch, the cause and the fault code
    _iStage := 0; _iReq := 0; // 作用域二：分级回零级 / scope two, the stage returns to zero
    _eState := E_DL_RagState.eNormal; // 作用域二：迁回正常相 / scope two, migrate to normal
    _fTprev := fTreactC; // 作用域三：温度快照重取（首拍不产生假速率）/ scope three, re-take the snapshot
    _fRateFilt := 0.0; // 作用域三：清速率滤波保持槽 / scope three, clear the rate filter hold slot
END_IF
// 段 4｜定时器与沿检测无条件周期刷新（R7），降级窗自复位（R188）
rtReset(CLK := bReset); // 复位沿无条件刷新 / unconditional refresh of the reset edge
tonDown(IN := (_iReq < _iStage) AND (NOT _bTrip) AND (NOT tonDown.Q), PT := _tDegrade); // 降级窗：需求低于当前级才计时，到期自复位 / the downgrade window with its own output inverted
// 段 5｜判据①温升速率：一阶差分 + 一阶指数滤波，分母零闸后计算（R4、R45 ②）
IF fDtSec > DL_RAG_DT_MIN THEN // 分母零闸 / the denominator gate
    _fRateRaw := (fTreactC - _fTprev) * DL_RAG_SEC_MIN / fDtSec; // 原始速率 [K/min] / the raw rate [K/min]
ELSE // 采样周期非法 / an illegal sample period
    _fRateRaw := 0.0; // 速率出零（不外推）/ the rate goes to zero
END_IF
IF NOT (_fRateRaw = _fRateRaw) THEN _fRateRaw := 0.0; END_IF // 速率 NaN 兜底 / the NaN fallback
IF (_fRateRaw - _fRateRaw) <> (_fRateRaw - _fRateRaw) THEN _fRateRaw := 0.0; END_IF // 速率 Inf 兜底 / the Inf fallback
_fTprev := fTreactC; // 上拍温度快照（差分用，用完立即赋值）/ the snapshot taken right after the difference
_fRateFilt := _fRateFilt + DL_RAG_RATE_ALPHA * (_fRateRaw - _fRateFilt); // 一阶指数滤波 [K/min] / the first order exponential filter [K/min]
IF NOT (_fRateFilt = _fRateFilt) THEN _fRateFilt := _fRateRaw; END_IF // 滤波结果 NaN 兜底 / the NaN fallback
IF (_fRateFilt - _fRateFilt) <> (_fRateFilt - _fRateFilt) THEN _fRateFilt := _fRateRaw; END_IF // 滤波结果 Inf 兜底 / the Inf fallback
// 段 6｜判据②绝热温升外推 MTSR：分母双零闸，外推上限兜底防发散（R4、R133）
IF (fBatchKg > DL_RAG_EPS) AND (fCpKjKgK > DL_RAG_EPS) THEN // 双分母零闸 / both denominators guarded
    _fFrac := fAccumKg / fBatchKg; // 已投料占比 [-] / the charged fraction [-]
    IF _fFrac < 0.0 THEN _fFrac := 0.0; ELSIF _fFrac > DL_RAG_FRAC_MAX THEN _fFrac := DL_RAG_FRAC_MAX; END_IF // 占比双向夹取 / clamp the fraction both ways
    _fMoles := fAccumKg / DL_RAG_MOLAR_KGKMOL; // 累积摩尔数 [kmol] / the accumulated moles [kmol]
    _fHeatKj := ABS(fDhKjMol) * DL_RAG_MOL_PER_KMOL * _fMoles; // 潜在放热量 [kJ] / the potential heat [kJ]
    _fDtAd := _fHeatKj / (fBatchKg * fCpKjKgK); // 绝热温升 [K] / the adiabatic rise [K]
    IF _fDtAd < 0.0 THEN _fDtAd := 0.0; ELSIF _fDtAd > DL_RAG_DTAD_MAX THEN _fDtAd := DL_RAG_DTAD_MAX; END_IF // 外推上限兜底 [K] / the extrapolation clamp [K]
ELSE // 组态越域 / the configuration is out of domain
    _fDtAd := 0.0; // 温升外推出零（不放大风险）/ the rise goes to zero and never inflates the risk
END_IF
_fMtsr := fTreactC + _fDtAd; // MTSR [°C] / the MTSR [°C]
// 段 7｜判据③冷却能力：温差与流量双源，温差反向加流量半限判完全失效
_fCoolDt := fTjacketC - fCoolInC; // 夹套与进水温差 [K] / the jacket to inlet difference [K]
_bCoolL5 := (_fCoolDt < 0.0) AND (fCoolFlowM3h < (fFlowMinM3h * DL_RAG_FLOW_L4_FRAC)); // 温差反向且流量低于半限＝冷却完全失效 / a reversed difference with less than half flow means no cooling
// 段 8｜三判据分档：逐判据独立档位与独立标志，成因不共用（R190）
_fRateThr1 := fRateTripKmin * DL_RAG_L1_FRAC; // 一档门限 [K/min] / the level one threshold [K/min]
_fRateThr2 := fRateTripKmin * DL_RAG_L2_FRAC; // 二档门限 [K/min] / the level two threshold [K/min]
_fRateThr3 := fRateTripKmin * DL_RAG_L3_FRAC; // 三档门限 [K/min] / the level three threshold [K/min]
_fRateThr4 := fRateTripKmin * DL_RAG_L4_FRAC; // 四档门限 [K/min] / the level four threshold [K/min]
_fMtsrThr1 := fMtsrLimitC - (fMtsrMarginK * DL_RAG_M1_FRAC); // 一档门限 [°C] / the level one threshold [°C]
_fMtsrThr2 := fMtsrLimitC - (fMtsrMarginK * DL_RAG_M2_FRAC); // 二档门限 [°C] / the level two threshold [°C]
_fMtsrThr3 := fMtsrLimitC - (fMtsrMarginK * DL_RAG_M3_FRAC); // 三档门限 [°C] / the level three threshold [°C]
_fMtsrThr4 := fMtsrLimitC - (fMtsrMarginK * DL_RAG_M4_FRAC); // 四档门限 [°C] / the level four threshold [°C]
_bRateL1 := _fRateFilt > _fRateThr1; // 判据①达一档 / criterion one at level one
_bRateL2 := _fRateFilt > _fRateThr2; // 判据①达二档 / criterion one at level two
_bRateL3 := _fRateFilt > _fRateThr3; // 判据①达三档 / criterion one at level three
_bRateL4 := _fRateFilt > _fRateThr4; // 判据①达四档 / criterion one at level four
_bRateL5 := _fRateFilt > fRateTripKmin; // 判据①达五档（独立成因标志）/ criterion one at level five
_iNeed := 0; // 判据①档位暂存清零 / clear the criterion one scratch
IF _bRateL5 THEN _iNeed := 5; ELSIF _bRateL4 THEN _iNeed := 4; ELSIF _bRateL3 THEN _iNeed := 3; ELSIF _bRateL2 THEN _iNeed := 2; ELSIF _bRateL1 THEN _iNeed := 1; END_IF // 判据①档位 / the criterion one level
IF _iNeed > _iReq THEN _iReq := _iNeed; END_IF // 合成取大 / aggregate by the maximum
_iNeed := 0; // 判据②档位暂存清零 / clear the criterion two scratch
IF _fMtsr > fMtsrLimitC THEN _iNeed := 5; // 判据②五档：超安全极限 / level five, the safety limit was passed
ELSIF _fMtsr > _fMtsrThr4 THEN _iNeed := 4; ELSIF _fMtsr > _fMtsrThr3 THEN _iNeed := 3; ELSIF _fMtsr > _fMtsrThr2 THEN _iNeed := 2; ELSIF _fMtsr > _fMtsrThr1 THEN _iNeed := 1; END_IF // 判据②一至四档 / the criterion two levels one to four
IF _iNeed > _iReq THEN _iReq := _iNeed; END_IF // 合成取大 / aggregate by the maximum
_iNeed := 0; // 判据③档位暂存清零 / clear the criterion three scratch
IF _bCoolL5 THEN // 冷却完全失效：直接五档（独立成因）/ a total cooling loss goes straight to level five
    _iNeed := 5; // 判据③五档 / criterion three at level five
ELSIF (_fCoolDt < 0.0) OR (fCoolFlowM3h < (fFlowMinM3h * DL_RAG_FLOW_L4_FRAC)) THEN // 温差反向或流量低于半限 / a reversed difference or less than half flow
    _iNeed := 4; // 判据③四档 / criterion three at level four
ELSIF (_fCoolDt < DL_RAG_COOL_DT_MIN) OR (fCoolFlowM3h < fFlowMinM3h) THEN // 温差不足或流量低于下限 / an insufficient difference or a flow below the floor
    _iNeed := 3; // 判据③三档 / criterion three at level three
END_IF
IF _iNeed > _iReq THEN _iReq := _iNeed; END_IF // 合成取大 / aggregate by the maximum
IF NOT xStirRun THEN // 搅拌停止：至少二级（独立于冷却与温度判据）/ a stopped agitator forces level two
    IF _iReq < 2 THEN _iReq := 2; END_IF // 二级下限 / the level two floor
END_IF
IF NOT bEnable THEN _iReq := 0; END_IF // 失能只清需求级，不解除全停锁存（R191 边界六）/ a disable clears the demand and never the latch
// 段 9｜故障锁存：每个成因独立枚举成员与独立码值，命中即置 bError 并同拍锁存（R45、R190）
IF NOT _bTrip THEN // 未锁存才判（锁存后一律回放，R152）/ judge only while unlatched
    IF NOT _bFinOk THEN // 入参非有限 / a non-finite input
        _eCause := E_DL_RagCause.eNotFinite; _iErrTmp := 2711; bError := TRUE; // 故障级成因、码位与标志（R45 配对）
    ELSIF NOT _bCfgOk THEN // 组态越域 / the configuration is out of domain
        _eCause := E_DL_RagCause.eCfgBad; _iErrTmp := 2712; bError := TRUE; // 故障级成因、码位与标志（R45 配对）
    ELSIF _bRateL5 THEN // 温升速率达五档 / the rate reached level five
        _eCause := E_DL_RagCause.eRateHigh; _iErrTmp := 2713; bError := TRUE; // 故障级成因、码位与标志（R45 配对）
    ELSIF _fMtsr > fMtsrLimitC THEN // MTSR 达五档 / the MTSR reached level five
        _eCause := E_DL_RagCause.eMtsrHigh; _iErrTmp := 2714; bError := TRUE; // 故障级成因、码位与标志（R45 配对）
    ELSIF _bCoolL5 THEN // 冷却完全失效 / the cooling was lost entirely
        _eCause := E_DL_RagCause.eCoolLoss; _iErrTmp := 2715; bError := TRUE; // 故障级成因、码位与标志（R45 配对）
    END_IF
    IF _iErrTmp <> 0 THEN // 存在故障级请求 / a fault grade request exists
        _iErrLch := _iErrTmp; _bTrip := TRUE; // 锁存码与锁存位单点写入 / the single write point of the code and the latch
    END_IF
END_IF
// 段 10｜分级仲裁：升级立即（安全侧优先）、降级按窗逐级（不跳级、不抖动）
IF _bTrip THEN // 已锁存 / already latched
    _iStage := 5; // 强制五级（锁存期内不降级）/ forced to level five while latched
ELSIF _iReq > _iStage THEN // 需求高于当前级：立即升级 / immediate escalation
    _iStage := _iReq; // 升级无延时（安全侧优先）/ escalation without delay
ELSIF (_iReq < _iStage) AND tonDown.Q THEN // 需求低于当前级且降级窗到期 / the demand is lower and the window expired
    _iStage := _iStage - 1; // 逐级降一级（每窗一级，禁跳级）/ one step per window
END_IF
IF _iStage < 0 THEN _iStage := 0; ELSIF _iStage > 5 THEN _iStage := 5; END_IF // 分级域夹取（防御性）/ clamp the stage domain
// 段 11｜相位映射：由分级单源映射、零滞后（R191），ELSE 落全停（R6）
CASE _iStage OF // 分级唯一权威 → 相位 / the single stage authority drives the phase
0: _eState := E_DL_RagState.eNormal; // 零级：正常 / level zero maps to normal
1: _eState := E_DL_RagState.eWarn; // 一级：报警 / level one maps to warn
2: _eState := E_DL_RagState.eStopFeed; // 二级：停止投料 / level two maps to stop feed
3: _eState := E_DL_RagState.eMaxCool; // 三级：加大冷却 / level three maps to maximum cooling
4: _eState := E_DL_RagState.eVent; // 四级：紧急泄放 / level four maps to venting
5: _eState := E_DL_RagState.eTrip; // 五级：全停 / level five maps to trip
ELSE // 非法分级值兜底（值域已夹取，防御性保留，R6、R128）
    _eState := E_DL_RagState.eTrip; // 落全停安全相 / fall back to the trip phase
    IF NOT _bTrip THEN // 未锁存才补锁存 / latch only while unlatched
        _eCause := E_DL_RagCause.eStageBad; _iErrLch := 2716; _bTrip := TRUE; bError := TRUE; // 故障级成因、码位与标志（R45 配对）
    END_IF
END_CASE
// 段 12｜统一出口：分级与五级位单源派生，连续量做非有限防护（R191、FB51-3）
iStage := _iStage; // 分级单点映射 / the single point mapping of the stage
xStage1 := _iStage >= 1; xStage2 := _iStage >= 2; xStage3 := _iStage >= 3; // 一至三级位（累积电平）/ levels one to three as accumulated levels
xStage4 := _iStage >= 4; xStage5 := _iStage >= 5; // 四至五级位（累积电平）/ levels four and five as accumulated levels
xAlarmOut := _iStage >= 1; xFeedStop := _iStage >= 2; xMaxCool := _iStage >= 3; // 一至三级动作输出 / the action outputs of levels one to three
xVentCmd := _iStage >= 4; xTotalStop := _iStage >= 5; // 四至五级动作输出 / the action outputs of levels four and five
xTripLatched := _bTrip; // 全停锁存回放 / replay the trip latch
eState := _eState; // 相位单点映射 / the single point mapping of the phase
fMtsrC := _fMtsr; // MTSR 单点映射 [°C] / the single point mapping of the MTSR [°C]
IF NOT (_fMtsr = _fMtsr) THEN fMtsrC := 0.0; END_IF // 出口 NaN 防护（安全侧出零）/ the NaN guard on the outlet
IF (_fMtsr - _fMtsr) <> (_fMtsr - _fMtsr) THEN fMtsrC := 0.0; END_IF // 出口 Inf 防护 / the Inf guard on the outlet
fRateKmin := _fRateFilt; // 速率单点映射 [K/min] / the single point mapping of the rate [K/min]
IF NOT (_fRateFilt = _fRateFilt) THEN fRateKmin := 0.0; END_IF // 出口 NaN 防护 / the NaN guard on the outlet
IF (_fRateFilt - _fRateFilt) <> (_fRateFilt - _fRateFilt) THEN fRateKmin := 0.0; END_IF // 出口 Inf 防护 / the Inf guard on the outlet
fDtAdK := _fDtAd; // 绝热温升单点映射 [K] / the single point mapping of the adiabatic rise [K]
xValid := _bFinOk AND _bCfgOk AND (NOT _bTrip); // 有效性：双闸通过且未锁存 / valid when both gates pass and nothing is latched
IF _bTrip THEN // 锁存期：故障级码回放，不按当下输入重推（R152）
    iErrCode := _iErrLch; bError := TRUE; // 锁存码回放、故障标志同源 / replay the code and share the latch source
ELSIF _iStage > 0 THEN // 未锁存但分级非零 / unlatched but a stage is active
    iErrCode := 2700 + _iStage; bError := FALSE; // 信息级动作码（每拍重算，不置故障标志，R45）/ the info action code without the fault flag
ELSE // 零级且未锁存 / level zero and unlatched
    iErrCode := 0; bError := FALSE; // 无码无标志 / no code and no flag
END_IF
END_FUNCTION_BLOCK

(* ---- FB_DL_ReactorYearWinClean.st ---- *)
(*==============================================================================
 * 组件名称 (Component)  : FB_DL_ReactorYearWinClean
 * 所属子库 (Sublibrary) : DL_Process
 * 当前版本 (Version)    : 1.0.0
 * 兼容性 (Platform)     : CODESYS 3.5+ / TwinCAT 3 / 汇川 InoProShop / 施耐德 Machine Expert
 *                         仅依赖 Standard.library（R_TRIG），零厂商私有库
 * 功能描述 (Function)   : 反应釜年度清洗窗与批次投料闸门。清洗窗内 CIP 完成
 *                         电平置「本窗已洗」锁存；窗内未洗或过窗未洗时投料
 *                         申请一律拒绝（批次闸门，拒绝成因独立分码 R190）；
 *                         窗关闭沿若整窗未洗 → bCleanOverdue 告警电平保持至
 *                         下窗。与 CipCleaningSeq（清洗执行顺控）分工：本件
 *                         职责在「门」不在「洗」——只判过窗未洗禁投料。
 * 来源标签 (Origin)     : ROADMAP §16.6 R11 池（L733），自研 clean-room
 * 边界语义 (Boundary)   : ① 「本窗已洗」锁存随窗开启沿清零（每窗独立判定）；
 *                         ② 窗电平输入为布尔域，无浮点量（无 NaN/除零域）；
 *                         ③ 窗内申请拒绝不锁存故障（业务拒绝态）；
 *                         ④ 过窗未洗告警清除路径 = 下窗开启沿或复位沿（头
 *                         注释声明）。
 * 输出语义 (Fallback)   : 【R191】bEnable = FALSE → 闸门出口强制 FALSE（拒绝
 *                         投料安全侧）；eFault 相 → 闸门 FALSE + bError。
 * 码位     (Codes)      : 按 R297 范式零 16# 码位硬编码；错误出口 BOOL+ENUM(eCause)。
 * 红线自检 (Redline)    : 7 项红线已自检：R1 零全局 ✓｜R2 零物理地址 ✓｜R3 纯 IEC ✓
 *                         R4 无浮点域 ✓｜R5 双语同行注释 ✓
 *                         R6 CASE 带 ELSE 兜底迁 eFault ✓｜R7 R_TRIG 段 0 无条件刷新 ✓
 * 验收向量 (Acceptance) : V1 窗内 + CIP 完成电平 → _bCleaned=TRUE，窗内申请
 *                         → bBatchAllow=TRUE；
 *                         V2 窗内未洗申请 → bBatchBlocked=TRUE，eDeny=eNotCleaned；
 *                         V3 窗关沿整窗未洗 → bCleanOverdue=TRUE 保持至下窗
 *                         开启沿清零。
 * 修订历史 (Revision)   : 2026-11-20  v1.0.0  R51 首版（批 2 · 序号 8）
 *==============================================================================*)
TYPE E_DL_RycDeny :
(
    eNone       := 0,                        (* 无拒绝（已放行或无申请） / No deny *)
    eNotCleaned := 1,                        (* 窗内未洗禁投 / Not cleaned this window *)
    eOverdue    := 2                         (* 过窗未洗禁投（告警期） / Overdue not cleaned *)
);
END_TYPE

TYPE E_DL_RycState :
(
    eIdle  := 0,                             (* 待使能 / Idle *)
    eGate  := 10,                            (* 闸门判定运行 / Gate run *)
    eFault := 90                             (* 故障锁存相 / Fault latched phase *)
);
END_TYPE

TYPE E_DL_RycCause :
(
    eNone     := 0,                          (* 无故障成因 / No cause *)
    ePhaseBad := 3                           (* 非法相位兜底 / Illegal phase fallback *)
);
END_TYPE

FUNCTION_BLOCK FB_DL_ReactorYearWinClean
VAR_INPUT
    bInCleanWin : BOOL := FALSE;             (* 年度清洗窗电平（上层窗判定供给）[-] / Clean-window level *)
    bCleanDone  : BOOL := FALSE;             (* CIP 清洗完成电平（CipCleaningSeq 供给）[-] / Clean-done level *)
    bBatchReq   : BOOL := FALSE;             (* 投料申请电平 [-] / Batch request *)
    bEnable     : BOOL := TRUE;              (* 使能 [-] / Enable *)
    bReset      : BOOL := FALSE;             (* 复位命令，上升沿清全部 [-] / Reset command *)
END_VAR
VAR_OUTPUT
    bBatchAllow  : BOOL;                     (* 投料放行电平（申请期实时）[-] / Batch allow level *)
    bBatchBlocked: BOOL;                     (* 投料拒绝电平（申请期实时）[-] / Batch blocked level *)
    eDeny        : E_DL_RycDeny;             (* 拒绝成因（信息级逐拍重算，R189） / Deny cause *)
    bCleanOverdue: BOOL;                     (* 过窗未洗告警电平（下窗开启沿或复位沿清，R152） / Overdue alarm *)
    nCleanWins   : UDINT;                    (* 累计完成清洗的窗数 [窗] / Cleaned window count *)
    eState       : E_DL_RycState;            (* 状态出口 / State outlet *)
    eCause       : E_DL_RycCause;            (* 故障成因出口 / Fault cause outlet *)
    bError       : BOOL;                     (* 故障锁存标志 [-] / Fault latch flag *)
END_VAR
VAR
    _eState    : E_DL_RycState := E_DL_RycState.eIdle;     (* 内部相位（CASE 唯一写入目标） / Internal phase *)
    _eCause    : E_DL_RycCause := E_DL_RycCause.eNone;     (* 故障成因锁存量 / Latched cause *)
    rtWinOpen  : R_TRIG;                     (* 窗开启沿实例，段 0 无条件调用 / Window-open edge *)
    rtWinClose : R_TRIG;                     (* 窗关闭沿实例，段 0 无条件调用 / Window-close edge *)
    rtReset    : R_TRIG;                     (* 复位沿实例，段 0 无条件调用 / Reset edge instance *)
    _bCleaned  : BOOL;                       (* 本窗已洗锁存 [-] / Cleaned-this-window latch *)
    _nWins     : UDINT;                      (* 完成清洗窗数锁存 [窗] / Cleaned-window count *)
    _bFault    : BOOL;                       (* 故障锁存位 / Latched fault bit *)
END_VAR

(* —— 段 0：沿实例无条件刷新（R228A；纯布尔域无浮点组态闸） —— *)
rtWinOpen(CLK := bInCleanWin);               (* 窗开启沿每拍必调 / Window-open edge every scan *)
rtWinClose(CLK := NOT bInCleanWin);          (* 窗关闭沿每拍必调 / Window-close edge every scan *)
rtReset(CLK := bReset);                      (* 复位沿每拍必调 / Reset edge every scan *)

(* —— 段 1：单拍量预清零（R107） —— *)
bBatchAllow := FALSE;                        (* 放行电平预清（判定分支覆盖） / Allow preset *)
bBatchBlocked := FALSE;                      (* 拒绝电平预清 / Blocked preset *)
eDeny := E_DL_RycDeny.eNone;                 (* 拒绝成因预清（信息级逐拍重算） / Deny preset *)

(* —— 段 2：复位沿处理（作用域：清故障 + 清已洗锁存 + 清告警 + 清窗数 + 迁 eIdle，R283 逐项声明） —— *)
IF rtReset.Q THEN
    _bFault := FALSE;                        (* 清故障锁存 / Clear fault *)
    _eCause := E_DL_RycCause.eNone;          (* 清成因 / Clear cause *)
    _bCleaned := FALSE;                      (* 清已洗锁存 / Clear cleaned latch *)
    bCleanOverdue := FALSE;                  (* 清过窗告警（复位沿清除路径之一，边界④） / Clear overdue *)
    _nWins := 0;                             (* 清窗数 / Clear count *)
    _eState := E_DL_RycState.eIdle;          (* 迁待机相 / Back to idle *)
END_IF

(* —— 段 4：CASE 主状态机（ELSE 兜底迁 eFault，红线 6） —— *)
CASE _eState OF
    E_DL_RycState.eIdle:                     (* 待机相 / Idle *)
        IF bEnable AND NOT _bFault THEN
            _eState := E_DL_RycState.eGate;  (* 进入闸门 / Enter gate *)
        END_IF
    E_DL_RycState.eGate:                     (* 闸门相：窗沿 + 已洗锁存 + 投料判定 / Gate *)
        IF NOT bEnable THEN
            _eState := E_DL_RycState.eIdle;  (* 失能回待机 / Back to idle *)
        ELSE
            IF rtWinOpen.Q THEN              (* 窗开启沿：本窗判定重置（边界①） + 上窗告警清除路径 / On window open *)
                _bCleaned := FALSE;          (* 清本窗已洗 / Reset cleaned latch *)
                bCleanOverdue := FALSE;      (* 清过窗告警（下窗开启沿清除路径，边界④） / Clear overdue *)
            END_IF
            IF bInCleanWin AND bCleanDone THEN
                _bCleaned := TRUE;           (* 窗内 CIP 完成：置已洗锁存（电平置位锁存语义） / Set cleaned latch *)
            END_IF
            IF rtWinClose.Q AND (NOT _bCleaned) THEN   (* 窗关沿整窗未洗：告警置位 / Overdue on close *)
                bCleanOverdue := TRUE;       (* 过窗未洗告警（保持至下窗/复位，R152） / Overdue alarm *)
            END_IF
            IF rtWinClose.Q AND _bCleaned THEN
                _nWins := _nWins + 1;        (* 完成清洗窗数（UDINT 回绕工程安全） / Count cleaned window *)
            END_IF
            IF bBatchReq THEN                (* 申请期实时判定（业务拒绝态不锁存故障，边界③） / On request *)
                IF bInCleanWin AND (NOT _bCleaned) THEN
                    bBatchBlocked := TRUE;   (* 窗内未洗拒绝 / Blocked *)
                    eDeny := E_DL_RycDeny.eNotCleaned;   (* 成因：未洗（独立成员，R190） / Cause: not cleaned *)
                ELSIF bCleanOverdue THEN
                    bBatchBlocked := TRUE;   (* 过窗未洗期拒绝 / Blocked *)
                    eDeny := E_DL_RycDeny.eOverdue;   (* 成因：过窗（独立成员） / Cause: overdue *)
                ELSE
                    bBatchAllow := TRUE;     (* 放行 / Allow *)
                END_IF
            END_IF
        END_IF
    E_DL_RycState.eFault:                    (* 故障相：冻结保持，仅复位沿出 / Fault *)
        ;                                    (* 锁存回放（R28） / Replay from latch *)
    ELSE                                     (* 非法相位兜底迁安全态 / Illegal phase fallback *)
        _eState := E_DL_RycState.eFault;     (* 迁故障相 / To fault *)
        _bFault := TRUE;                     (* 同步锁存 / Latch *)
        _eCause := E_DL_RycCause.ePhaseBad;  (* 成因：非法相位 / Cause: illegal phase *)
END_CASE

(* —— 段 5：出口映射（bError/eState 同源，R191） —— *)
nCleanWins := _nWins;                        (* 窗数出口 / Count outlet *)
bError := _bFault;                           (* 故障标志镜像 / Fault flag mirror *)
eState := _eState;                           (* 状态出口 / State outlet *)
eCause := _eCause;                           (* 成因出口 / Cause outlet *)
END_FUNCTION_BLOCK

(* ---- FB_DL_RecipeSearchFifo.st ---- *)
(*
  FB_DL_RecipeSearchFifo  —  配方请求 FIFO 排队（队列 + 校验链） / Recipe request FIFO queue with checksum chain
  分类 Category : DL_Process
  版本 Version  : 1.0.0
  来源 Source   : t1-4-codesys-forge — 队列/调度族零检索深化（与 RecipeManager 配方主件分工：那件管配方存取，本件管请求排队）
  溯源 Origin   : clean-room 实现，未复制任何源码行
  功能 Function : 1) 深度 8 固定 FIFO：bEnqCmd 沿入队（uReqId 入栈，异或校验链
                  uChecksum := uReqId XOR 16#A5A5_A5A5 入栈承载），bDeqCmd 沿
                  出队并校验链复核（uReqId XOR 16#A5A5_A5A5 = uChecksum 才放行）；
                  2) 故障级三码独立：038B 队满入队拒收锁存 / 038C 出队校验链
                  失败锁存（数据完整性违约，R190 归因唯一）/ 038D 空队出队违约
                  锁存 + ELSE 兜底归并（码表声明）；
                  3) 信息级三码：入队成功 / 出队成功 / 校验链复核通过（单拍沿）；
                  4) 首尾游标 MOD 8 回绕（除数 8 为常量无除零），计满/排空两端
                  边界即整数进位点验收向量（R28-2：count=8 与 count=0 两点）；
                  5) 解除式全当拍量（R240 落地），逐 BOOL 标注见段 4。
  边界 Boundary : ① 游标域 0..7 由常量 8 的 MOD 结构性限定，无越界路径；
                  ② 队列内容快照仅在命令沿承载（锁存量），每拍不重扫；
                  ③ 校验链为完整性哨兵非加密（头注释声明，防误读）；
                  ④ 无 GVL 依赖：纯引脚输入输出，无外部变量引用，无物理 IO 地址。
  依赖 Depends  : Standard.library（R_TRIG）
  码表 Error codes（Process 段 0005，窗口 038B~038D / 04B3~04B5）:
    16#0005_038B 故障级：队满入队拒收锁存（count = 8 仍入队），锁存至 bReset
    16#0005_038C 故障级：出队校验链失败锁存（异或复核不匹配），锁存至 bReset
    16#0005_038D 故障级：空队出队违约或相位落 ELSE 兜底（归并声明），锁存至 bReset
    16#0005_04B3 信息级：入队成功沿
    16#0005_04B4 信息级：出队成功沿
    16#0005_04B5 信息级：出队校验链复核通过沿
  修订历史 Revision :
    2026-11-19  v1.0.0  R42 首版（批次 2 · 序号 5）
*)

TYPE ST_DL_RqEntry :
STRUCT
    uReqId    : UDINT;              // 请求配方号 [-] / Requested recipe ID
    uChecksum : UDINT;              // 入队校验链（uReqId 异或哨兵）[-] / Enqueue checksum chain
END_STRUCT
END_TYPE

TYPE E_DL_RsfState :
(
    eIdle   := 0,    // 空闲：队列待命 / Idle, queue standing by
    eFault  := 90    // 故障：契约违约锁定 / Fault, latched
);
END_TYPE

FUNCTION_BLOCK FB_DL_RecipeSearchFifo
VAR_INPUT
    bEnqCmd      : BOOL := FALSE;     // 入队命令，上升沿承载 [-] / Enqueue command edge
    uReqId       : UDINT := 0;        // 入队请求配方号（bEnqCmd 沿采信）[-] / Enqueue recipe ID
    bDeqCmd      : BOOL := FALSE;     // 出队命令，上升沿承载 [-] / Dequeue command edge
    bReset       : BOOL := FALSE;     // 复位，上升沿清故障锁存与队列 / Reset edge clears fault and queue
END_VAR
VAR_OUTPUT
    eState       : E_DL_RsfState;     // 状态出口，段尾单点映射 / State outlet
    nCount       : DINT;              // 当前队列深度 [0..8] / Current queue depth
    uDeqId       : UDINT;             // 出队配方号（校验通过后有效）[-] / Dequeued recipe ID
    bDeqValid    : BOOL;              // 出队有效单拍镜像 [-] / Dequeue valid one-shot mirror
    bQueueFull   : BOOL;              // 队满镜像（count = 8）[-] / Queue-full mirror
    bError       : BOOL;              // 故障锁存标志 / Fault latch flag
    nErrId       : UDINT;             // 事件码，0 = 无事件 / Event code
END_VAR
VAR
    a_stQueue    : ARRAY[0..7] OF ST_DL_RqEntry;  // 8 深度队列存储 / Queue storage
    rtEnq        : R_TRIG;            // 入队沿实例，无条件刷新 / Enqueue edge instance
    rtDeq        : R_TRIG;            // 出队沿实例，无条件刷新 / Dequeue edge instance
    rtReset      : R_TRIG;            // 复位沿实例，无条件刷新 / Reset edge instance
    _nHead       : DINT := 0;         // 队头游标 [0..7]（出队位置）/ Head cursor
    _nTail       : DINT := 0;         // 队尾游标 [0..7]（入队位置）/ Tail cursor
    _nCnt        : DINT := 0;         // 队列深度计数 [0..8] / Depth counter
    _bFault      : BOOL;              // 故障锁存位（锁存量）/ Latched fault bit
    _eState      : E_DL_RsfState := E_DL_RsfState.eIdle;   // 内部相位，段 5A 唯一写入目标 / Internal phase, the only write target of segment 5A
    _uFault      : UDINT;             // 故障码锁存（锁存量）/ Latched fault code
    _uInfo       : UDINT;             // 信息码，每拍重算 / Transient info code
END_VAR

(* —— 段 0：沿实例无条件周期刷新（禁置于 IF/CASE 内） —— *)
rtEnq(CLK := bEnqCmd);               // 入队沿（每拍必调）
rtDeq(CLK := bDeqCmd);               // 出队沿（每拍必调）
rtReset(CLK := bReset);              // 复位沿（每拍必调）

(* —— 段 1：单拍量预清零（锁存量 _bFault/_uFault 与游标/队列不入清单，禁同拍抹除） —— *)
_uInfo := 16#0000_0000;             // 信息码每拍重算
bDeqValid := FALSE;                 // 出队有效镜像缺省 FALSE（单拍）
uDeqId := 16#0000_0000;             // 出队号缺省 0
nErrId := 16#0000_0000;             // 事件码缺省无事件

(* —— 段 2：复位沿（判据当拍量；清锁存与全队列） —— *)
IF rtReset.Q THEN                   // rtReset.Q = 当拍量
    _bFault := FALSE;               // 清故障锁存位
    _uFault := 16#0000_0000;        // 清故障锁存码
    _nHead := 0;                    // 队头游标清零
    _nTail := 0;                    // 队尾游标清零
    _nCnt := 0;                     // 深度计数清零
END_IF

(* —— 段 3：入队承载（判据当拍量沿；count = 8 满界为进位点验收向量之一） —— *)
IF rtEnq.Q AND (NOT _bFault) THEN
    IF _nCnt >= 8 THEN              // 队满（上界进位点）
        _uFault := 16#0005_038B;    // 故障级：队满入队拒收
        _bFault := TRUE;            // 故障标志与码位配对（R45）
    ELSE
        a_stQueue[_nTail].uReqId := uReqId;             // 请求号入栈
        a_stQueue[_nTail].uChecksum := uReqId XOR 16#A5A5_A5A5;  // 校验链入栈（异或哨兵）
        _nTail := (_nTail + 1) MOD 8;                   // 队尾游标回绕（除数 8 常量无除零）
        _nCnt := _nCnt + 1;                             // 深度递增
        _uInfo := 16#0005_04B3;         // 信息级：入队成功沿
    END_IF
END_IF

(* —— 段 4：出队承载（判据当拍量沿；count = 0 空界为进位点验收向量之一） —— *)
IF rtDeq.Q AND (NOT _bFault) THEN
    IF _nCnt = 0 THEN               // 空队（下界进位点）
        _uFault := 16#0005_038D;    // 故障级：空队出队违约
        _bFault := TRUE;
    ELSE
        IF (a_stQueue[_nHead].uReqId XOR 16#A5A5_A5A5) = a_stQueue[_nHead].uChecksum THEN
            uDeqId := a_stQueue[_nHead].uReqId;         // 校验通过：出队号放行
            bDeqValid := TRUE;      // 出队有效单拍镜像
            _uInfo := 16#0005_04B5; // 信息级：校验链复核通过沿
        ELSE
            _uFault := 16#0005_038C;    // 故障级：校验链失败（数据完整性违约）
            _bFault := TRUE;
        END_IF
        _nHead := (_nHead + 1) MOD 8;                   // 队头游标回绕（除数 8 常量）
        IF NOT _bFault THEN
            _nCnt := _nCnt - 1;     // 深度递减（校验失败拍不递减，保现场）
            _uInfo := 16#0005_04B4; // 信息级：出队成功沿（覆盖通过沿，后到优先声明）
        END_IF
    END_IF
END_IF

(* —— 段 5：故障解除式（R240 落地，逐 BOOL 标注）：
     rtReset.Q = 当拍量；NOT bEnqCmd = 当拍量；NOT bDeqCmd = 当拍量。
     均不含锁存量（_bFault/_uFault），解除边真实可达（命令撤销 + 复位沿）。 —— *)
IF rtReset.Q AND (NOT bEnqCmd) AND (NOT bDeqCmd) THEN
    _bFault := FALSE;               // 清故障锁存位（锁存量，仅此当拍量解除沿可清）
    _uFault := 16#0000_0000;        // 清故障锁存码（锁存量，仅本当拍量解除沿可清）
END_IF

(* —— 段 5A：状态相位更新（_eState 唯一写入目标，与锁存位同源） —— *)
IF _bFault THEN
    _eState := E_DL_RsfState.eFault;    // 故障锁存即入故障相 / Fault latch enters fault phase
ELSE
    _eState := E_DL_RsfState.eIdle;     // 非故障为空闲待命相 / Non-fault is the idle phase
END_IF

(* —— 段 6：出口单点映射（名实同源；锁存码回放，禁同拍抹除） —— *)
IF _bFault THEN
    nErrId := _uFault;              // 故障锁存码回放
    bDeqValid := FALSE;             // 故障拍出队有效镜像强制 FALSE（安全侧）
ELSE
    nErrId := _uInfo;               // 信息码
END_IF
nCount := _nCnt;                    // 深度出口
bQueueFull := (_nCnt >= 8);         // 队满镜像（上界进位点直读）
bError := _bFault;                  // 故障标志与锁存位同源
eState := _eState;                  // 状态出口单点映射

END_FUNCTION_BLOCK
